    ELSIF ((x0 = TRUE) AND  (t0.Q = TRUE) AND  (t1.Q = FALSE)) THEN 
        cstate16 := 38115; y0 := TRUE; y1 := FALSE; y2 := FALSE; t0_start := TRUE; t0_up := FALSE;t1_start := FALSE; 
    ELSIF ((x0 = TRUE) AND  (t0.Q = TRUE) AND  (t1.Q = TRUE)) THEN 
        cstate16 := 39140; y0 := TRUE; y1 := FALSE; y2 := FALSE; t0_start := TRUE; t0_up := FALSE;t1_start := FALSE; 
    END_IF;
42457:
    IF ((x0 = FALSE) AND  (t0.Q = FALSE) AND  (t1.Q = FALSE)) THEN 
        cstate16 := 32883; y0 := FALSE; y1 := FALSE; y2 := FALSE; t0_start := FALSE;t1_start := FALSE; 
    ELSIF ((x0 = FALSE) AND  (t0.Q = FALSE) AND  (t1.Q = TRUE)) THEN 
        cstate16 := 34932; y0 := FALSE; y1 := FALSE; y2 := FALSE; t0_start := FALSE;t1_start := FALSE; 
    ELSIF ((x0 = FALSE) AND  (t0.Q = TRUE) AND  (t1.Q = FALSE)) THEN 
        cstate16 := 27763; y0 := FALSE; y1 := FALSE; y2 := FALSE; t0_start := FALSE;t1_start := FALSE; 
    ELSIF ((x0 = FALSE) AND  (t0.Q = TRUE) AND  (t1.Q = TRUE)) THEN 
        cstate16 := 28788; y0 := FALSE; y1 := FALSE; y2 := FALSE; t0_start := FALSE;t1_start := FALSE; 
    ELSIF ((x0 = TRUE) AND  (t0.Q = FALSE) AND  (t1.Q = FALSE)) THEN 
        cstate16 := 49657; y0 := TRUE; y1 := TRUE; y2 := TRUE; t0_start := FALSE;t1_start := FALSE; 
    ELSIF ((x0 = TRUE) AND  (t0.Q = FALSE) AND  (t1.Q = TRUE)) THEN 
        cstate16 := 48646; y0 := TRUE; y1 := TRUE; y2 := TRUE; t0_start := FALSE;t1_start := FALSE; 
    ELSIF ((x0 = TRUE) AND  (t0.Q = TRUE) AND  (t1.Q = FALSE)) THEN 
        cstate16 := 42489; y0 := TRUE; y1 := TRUE; y2 := TRUE; t0_start := FALSE;t1_start := FALSE; 
    ELSIF ((x0 = TRUE) AND  (t0.Q = TRUE) AND  (t1.Q = TRUE)) THEN 
        cstate16 := 43526; y0 := TRUE; y1 := TRUE; y2 := TRUE; t0_start := FALSE;t1_start := FALSE; 
    END_IF;
27731:
    IF ((x0 = FALSE) AND  (t0.Q = FALSE) AND  (t1.Q = FALSE)) THEN 
        cstate16 := 32883; y0 := FALSE; y1 := FALSE; y2 := FALSE; t0_start := FALSE;t1_start := FALSE; 
    ELSIF ((x0 = FALSE) AND  (t0.Q = FALSE) AND  (t1.Q = TRUE)) THEN 
        cstate16 := 34932; y0 := FALSE; y1 := FALSE; y2 := FALSE; t0_start := FALSE;t1_start := FALSE; 
    ELSIF ((x0 = FALSE) AND  (t0.Q = TRUE) AND  (t1.Q = FALSE)) THEN 
        cstate16 := 27763; y0 := FALSE; y1 := FALSE; y2 := FALSE; t0_start := FALSE;t1_start := FALSE; 
    ELSIF ((x0 = FALSE) AND  (t0.Q = TRUE) AND  (t1.Q = TRUE)) THEN 
        cstate16 := 28788; y0 := FALSE; y1 := FALSE; y2 := FALSE; t0_start := FALSE;t1_start := FALSE; 
    ELSIF ((x0 = TRUE) AND  (t0.Q = FALSE) AND  (t1.Q = FALSE)) THEN 
        cstate16 := 41187; y0 := TRUE; y1 := FALSE; y2 := FALSE; t0_start := TRUE; t0_up := FALSE;t1_start := FALSE; 
    ELSIF ((x0 = TRUE) AND  (t0.Q = FALSE) AND  (t1.Q = TRUE)) THEN 
        cstate16 := 40167; y0 := TRUE; y1 := FALSE; y2 := TRUE; t0_start := TRUE; t0_up := FALSE;t1_start := FALSE; 
    ELSIF ((x0 = TRUE) AND  (t0.Q = TRUE) AND  (t1.Q = FALSE)) THEN 
        cstate16 := 38115; y0 := TRUE; y1 := FALSE; y2 := FALSE; t0_start := TRUE; t0_up := FALSE;t1_start := FALSE; 
    ELSIF ((x0 = TRUE) AND  (t0.Q = TRUE) AND  (t1.Q = TRUE)) THEN 
        cstate16 := 39143; y0 := TRUE; y1 := FALSE; y2 := TRUE; t0_start := TRUE; t0_up := FALSE;t1_start := FALSE; 
    END_IF;
41555:
    IF ((x0 = FALSE) AND  (t0.Q = FALSE) AND  (t1.Q = FALSE)) THEN 
        cstate16 := 23667; y0 := FALSE; y1 := FALSE; y2 := FALSE; t0_start := FALSE;t1_start := FALSE; 
    ELSIF ((x0 = FALSE) AND  (t0.Q = FALSE) AND  (t1.Q = TRUE)) THEN 
        cstate16 := 26740; y0 := FALSE; y1 := FALSE; y2 := FALSE; t0_start := FALSE;t1_start := FALSE; 
    ELSIF ((x0 = FALSE) AND  (t0.Q = TRUE) AND  (t1.Q = FALSE)) THEN 
        cstate16 := 17491; y0 := FALSE; y1 := FALSE; y2 := FALSE; t0_start := FALSE;t1_start := TRUE; t1_up := FALSE; 
    ELSIF ((x0 = FALSE) AND  (t0.Q = TRUE) AND  (t1.Q = TRUE)) THEN 
        cstate16 := 17492; y0 := FALSE; y1 := FALSE; y2 := FALSE; t0_start := FALSE;t1_start := TRUE; t1_up := FALSE; 
    ELSIF ((x0 = TRUE) AND  (t0.Q = FALSE) AND  (t1.Q = FALSE)) THEN 
        cstate16 := 41555; y0 := TRUE; y1 := FALSE; y2 := FALSE; t0_start := FALSE;t1_start := FALSE; 
    ELSIF ((x0 = TRUE) AND  (t0.Q = FALSE) AND  (t1.Q = TRUE)) THEN 
        cstate16 := 40535; y0 := TRUE; y1 := FALSE; y2 := TRUE; t0_start := FALSE;t1_start := FALSE; 
    ELSIF ((x0 = TRUE) AND  (t0.Q = TRUE) AND  (t1.Q = FALSE)) THEN 
        cstate16 := 46643; y0 := TRUE; y1 := TRUE; y2 := FALSE; t0_start := FALSE;t1_start := TRUE; t1_up := FALSE; 
    ELSIF ((x0 = TRUE) AND  (t0.Q = TRUE) AND  (t1.Q = TRUE)) THEN 
        cstate16 := 46648; y0 := TRUE; y1 := TRUE; y2 := TRUE; t0_start := FALSE;t1_start := TRUE; t1_up := FALSE; 
    END_IF;
42453:
    IF ((x0 = FALSE) AND  (t0.Q = FALSE) AND  (t1.Q = FALSE)) THEN 
        cstate16 := 32883; y0 := FALSE; y1 := FALSE; y2 := FALSE; t0_start := FALSE;t1_start := FALSE; 
    ELSIF ((x0 = FALSE) AND  (t0.Q = FALSE) AND  (t1.Q = TRUE)) THEN 
        cstate16 := 34932; y0 := FALSE; y1 := FALSE; y2 := FALSE; t0_start := FALSE;t1_start := FALSE; 
    ELSIF ((x0 = FALSE) AND  (t0.Q = TRUE) AND  (t1.Q = FALSE)) THEN 
        cstate16 := 27763; y0 := FALSE; y1 := FALSE; y2 := FALSE; t0_start := FALSE;t1_start := FALSE; 
    ELSIF ((x0 = FALSE) AND  (t0.Q = TRUE) AND  (t1.Q = TRUE)) THEN 
        cstate16 := 28788; y0 := FALSE; y1 := FALSE; y2 := FALSE; t0_start := FALSE;t1_start := FALSE; 
    ELSIF ((x0 = TRUE) AND  (t0.Q = FALSE) AND  (t1.Q = FALSE)) THEN 
        cstate16 := 49657; y0 := TRUE; y1 := TRUE; y2 := TRUE; t0_start := FALSE;t1_start := FALSE; 
    ELSIF ((x0 = TRUE) AND  (t0.Q = FALSE) AND  (t1.Q = TRUE)) THEN 
        cstate16 := 48646; y0 := TRUE; y1 := TRUE; y2 := TRUE; t0_start := FALSE;t1_start := FALSE; 
    ELSIF ((x0 = TRUE) AND  (t0.Q = TRUE) AND  (t1.Q = FALSE)) THEN 
        cstate16 := 42489; y0 := TRUE; y1 := TRUE; y2 := TRUE; t0_start := FALSE;t1_start := FALSE; 
    ELSIF ((x0 = TRUE) AND  (t0.Q = TRUE) AND  (t1.Q = TRUE)) THEN 
        cstate16 := 43526; y0 := TRUE; y1 := TRUE; y2 := TRUE; t0_start := FALSE;t1_start := FALSE; 
    END_IF;
42450:
    IF ((x0 = FALSE) AND  (t0.Q = FALSE) AND  (t1.Q = FALSE)) THEN 
        cstate16 := 32883; y0 := FALSE; y1 := FALSE; y2 := FALSE; t0_start := FALSE;t1_start := FALSE; 
    ELSIF ((x0 = FALSE) AND  (t0.Q = FALSE) AND  (t1.Q = TRUE)) THEN 
        cstate16 := 34932; y0 := FALSE; y1 := FALSE; y2 := FALSE; t0_start := FALSE;t1_start := FALSE; 
    ELSIF ((x0 = FALSE) AND  (t0.Q = TRUE) AND  (t1.Q = FALSE)) THEN 
        cstate16 := 27763; y0 := FALSE; y1 := FALSE; y2 := FALSE; t0_start := FALSE;t1_start := FALSE; 
    ELSIF ((x0 = FALSE) AND  (t0.Q = TRUE) AND  (t1.Q = TRUE)) THEN 
        cstate16 := 28788; y0 := FALSE; y1 := FALSE; y2 := FALSE; t0_start := FALSE;t1_start := FALSE; 
    ELSIF ((x0 = TRUE) AND  (t0.Q = FALSE) AND  (t1.Q = FALSE)) THEN 
        cstate16 := 49649; y0 := TRUE; y1 := TRUE; y2 := FALSE; t0_start := FALSE;t1_start := FALSE; 
    ELSIF ((x0 = TRUE) AND  (t0.Q = FALSE) AND  (t1.Q = TRUE)) THEN 
        cstate16 := 48642; y0 := TRUE; y1 := TRUE; y2 := FALSE; t0_start := FALSE;t1_start := FALSE; 
    ELSIF ((x0 = TRUE) AND  (t0.Q = TRUE) AND  (t1.Q = FALSE)) THEN 
        cstate16 := 42481; y0 := TRUE; y1 := TRUE; y2 := FALSE; t0_start := FALSE;t1_start := FALSE; 
    ELSIF ((x0 = TRUE) AND  (t0.Q = TRUE) AND  (t1.Q = TRUE)) THEN 
        cstate16 := 43522; y0 := TRUE; y1 := TRUE; y2 := FALSE; t0_start := FALSE;t1_start := FALSE; 
    END_IF;
26740:
    IF ((x0 = FALSE) AND  (t0.Q = FALSE) AND  (t1.Q = FALSE)) THEN 
        cstate16 := 26739; y0 := FALSE; y1 := FALSE; y2 := FALSE; t0_start := FALSE;t1_start := FALSE; 
    ELSIF ((x0 = FALSE) AND  (t0.Q = FALSE) AND  (t1.Q = TRUE)) THEN 
        cstate16 := 26740; y0 := FALSE; y1 := FALSE; y2 := FALSE; t0_start := FALSE;t1_start := FALSE; 
    ELSIF ((x0 = FALSE) AND  (t0.Q = TRUE) AND  (t1.Q = FALSE)) THEN 
        cstate16 := 17491; y0 := FALSE; y1 := FALSE; y2 := FALSE; t0_start := FALSE;t1_start := TRUE; t1_up := FALSE; 
    ELSIF ((x0 = FALSE) AND  (t0.Q = TRUE) AND  (t1.Q = TRUE)) THEN 
        cstate16 := 17492; y0 := FALSE; y1 := FALSE; y2 := FALSE; t0_start := FALSE;t1_start := TRUE; t1_up := FALSE; 
    ELSIF ((x0 = TRUE) AND  (t0.Q = FALSE) AND  (t1.Q = FALSE)) THEN 
        cstate16 := 40163; y0 := TRUE; y1 := FALSE; y2 := FALSE; t0_start := TRUE; t0_up := FALSE;t1_start := FALSE; 
    ELSIF ((x0 = TRUE) AND  (t0.Q = FALSE) AND  (t1.Q = TRUE)) THEN 
        cstate16 := 40164; y0 := TRUE; y1 := FALSE; y2 := FALSE; t0_start := TRUE; t0_up := FALSE;t1_start := FALSE; 
    ELSIF ((x0 = TRUE) AND  (t0.Q = TRUE) AND  (t1.Q = FALSE)) THEN 
        cstate16 := 38147; y0 := TRUE; y1 := TRUE; y2 := FALSE; t0_start := TRUE; t0_up := FALSE;t1_start := TRUE; t1_up := FALSE; 
    ELSIF ((x0 = TRUE) AND  (t0.Q = TRUE) AND  (t1.Q = TRUE)) THEN 
        cstate16 := 38148; y0 := TRUE; y1 := TRUE; y2 := FALSE; t0_start := TRUE; t0_up := FALSE;t1_start := TRUE; t1_up := FALSE; 
    END_IF;
40532:
    IF ((x0 = FALSE) AND  (t0.Q = FALSE) AND  (t1.Q = FALSE)) THEN 
        cstate16 := 26739; y0 := FALSE; y1 := FALSE; y2 := FALSE; t0_start := FALSE;t1_start := FALSE; 
    ELSIF ((x0 = FALSE) AND  (t0.Q = FALSE) AND  (t1.Q = TRUE)) THEN 
        cstate16 := 26740; y0 := FALSE; y1 := FALSE; y2 := FALSE; t0_start := FALSE;t1_start := FALSE; 
    ELSIF ((x0 = FALSE) AND  (t0.Q = TRUE) AND  (t1.Q = FALSE)) THEN 
        cstate16 := 17491; y0 := FALSE; y1 := FALSE; y2 := FALSE; t0_start := FALSE;t1_start := TRUE; t1_up := FALSE; 
    ELSIF ((x0 = FALSE) AND  (t0.Q = TRUE) AND  (t1.Q = TRUE)) THEN 
        cstate16 := 17492; y0 := FALSE; y1 := FALSE; y2 := FALSE; t0_start := FALSE;t1_start := TRUE; t1_up := FALSE; 
    ELSIF ((x0 = TRUE) AND  (t0.Q = FALSE) AND  (t1.Q = FALSE)) THEN 
        cstate16 := 40531; y0 := TRUE; y1 := FALSE; y2 := FALSE; t0_start := FALSE;t1_start := FALSE; 
    ELSIF ((x0 = TRUE) AND  (t0.Q = FALSE) AND  (t1.Q = TRUE)) THEN 
        cstate16 := 40532; y0 := TRUE; y1 := FALSE; y2 := FALSE; t0_start := FALSE;t1_start := FALSE; 
    ELSIF ((x0 = TRUE) AND  (t0.Q = TRUE) AND  (t1.Q = FALSE)) THEN 
        cstate16 := 46643; y0 := TRUE; y1 := TRUE; y2 := FALSE; t0_start := FALSE;t1_start := TRUE; t1_up := FALSE; 
    ELSIF ((x0 = TRUE) AND  (t0.Q = TRUE) AND  (t1.Q = TRUE)) THEN 
        cstate16 := 46644; y0 := TRUE; y1 := TRUE; y2 := FALSE; t0_start := FALSE;t1_start := TRUE; t1_up := FALSE; 
    END_IF;
40535:
    IF ((x0 = FALSE) AND  (t0.Q = FALSE) AND  (t1.Q = FALSE)) THEN 
        cstate16 := 26739; y0 := FALSE; y1 := FALSE; y2 := FALSE; t0_start := FALSE;t1_start := FALSE; 
    ELSIF ((x0 = FALSE) AND  (t0.Q = FALSE) AND  (t1.Q = TRUE)) THEN 
        cstate16 := 26740; y0 := FALSE; y1 := FALSE; y2 := FALSE; t0_start := FALSE;t1_start := FALSE; 
    ELSIF ((x0 = FALSE) AND  (t0.Q = TRUE) AND  (t1.Q = FALSE)) THEN 
        cstate16 := 17491; y0 := FALSE; y1 := FALSE; y2 := FALSE; t0_start := FALSE;t1_start := TRUE; t1_up := FALSE; 
    ELSIF ((x0 = FALSE) AND  (t0.Q = TRUE) AND  (t1.Q = TRUE)) THEN 
        cstate16 := 17492; y0 := FALSE; y1 := FALSE; y2 := FALSE; t0_start := FALSE;t1_start := TRUE; t1_up := FALSE; 
    ELSIF ((x0 = TRUE) AND  (t0.Q = FALSE) AND  (t1.Q = FALSE)) THEN 
        cstate16 := 40540; y0 := TRUE; y1 := FALSE; y2 := TRUE; t0_start := FALSE;t1_start := FALSE; 
    ELSIF ((x0 = TRUE) AND  (t0.Q = FALSE) AND  (t1.Q = TRUE)) THEN 
        cstate16 := 40535; y0 := TRUE; y1 := FALSE; y2 := TRUE; t0_start := FALSE;t1_start := FALSE; 
    ELSIF ((x0 = TRUE) AND  (t0.Q = TRUE) AND  (t1.Q = FALSE)) THEN 
        cstate16 := 46651; y0 := TRUE; y1 := TRUE; y2 := TRUE; t0_start := FALSE;t1_start := TRUE; t1_up := FALSE; 
    ELSIF ((x0 = TRUE) AND  (t0.Q = TRUE) AND  (t1.Q = TRUE)) THEN 
        cstate16 := 46648; y0 := TRUE; y1 := TRUE; y2 := TRUE; t0_start := FALSE;t1_start := TRUE; t1_up := FALSE; 
    END_IF;
6481:
    IF ((x0 = FALSE) AND  (t0.Q = FALSE) AND  (t1.Q = FALSE)) THEN 
        cstate16 := 34931; y0 := FALSE; y1 := FALSE; y2 := FALSE; t0_start := FALSE;t1_start := FALSE; 
    ELSIF ((x0 = FALSE) AND  (t0.Q = FALSE) AND  (t1.Q = TRUE)) THEN 
        cstate16 := 34932; y0 := FALSE; y1 := FALSE; y2 := FALSE; t0_start := FALSE;t1_start := FALSE; 
    ELSIF ((x0 = FALSE) AND  (t0.Q = TRUE) AND  (t1.Q = FALSE)) THEN 
        cstate16 := 28787; y0 := FALSE; y1 := FALSE; y2 := FALSE; t0_start := FALSE;t1_start := FALSE; 
    ELSIF ((x0 = FALSE) AND  (t0.Q = TRUE) AND  (t1.Q = TRUE)) THEN 
        cstate16 := 28788; y0 := FALSE; y1 := FALSE; y2 := FALSE; t0_start := FALSE;t1_start := FALSE; 
    ELSIF ((x0 = TRUE) AND  (t0.Q = FALSE) AND  (t1.Q = FALSE)) THEN 
        cstate16 := 14673; y0 := FALSE; y1 := TRUE; y2 := FALSE; t0_start := FALSE;t1_start := FALSE; 
    ELSIF ((x0 = TRUE) AND  (t0.Q = FALSE) AND  (t1.Q = TRUE)) THEN 
        cstate16 := 14678; y0 := FALSE; y1 := TRUE; y2 := TRUE; t0_start := FALSE;t1_start := FALSE; 
    ELSIF ((x0 = TRUE) AND  (t0.Q = TRUE) AND  (t1.Q = FALSE)) THEN 
        cstate16 := 6481; y0 := FALSE; y1 := TRUE; y2 := FALSE; t0_start := FALSE;t1_start := FALSE; 
    ELSIF ((x0 = TRUE) AND  (t0.Q = TRUE) AND  (t1.Q = TRUE)) THEN 
        cstate16 := 6486; y0 := FALSE; y1 := TRUE; y2 := TRUE; t0_start := FALSE;t1_start := FALSE; 
    END_IF;
6482:
    IF ((x0 = FALSE) AND  (t0.Q = FALSE) AND  (t1.Q = FALSE)) THEN 
        cstate16 := 34931; y0 := FALSE; y1 := FALSE; y2 := FALSE; t0_start := FALSE;t1_start := FALSE; 
    ELSIF ((x0 = FALSE) AND  (t0.Q = FALSE) AND  (t1.Q = TRUE)) THEN 
        cstate16 := 34932; y0 := FALSE; y1 := FALSE; y2 := FALSE; t0_start := FALSE;t1_start := FALSE; 
    ELSIF ((x0 = FALSE) AND  (t0.Q = TRUE) AND  (t1.Q = FALSE)) THEN 
        cstate16 := 28787; y0 := FALSE; y1 := FALSE; y2 := FALSE; t0_start := FALSE;t1_start := FALSE; 
    ELSIF ((x0 = FALSE) AND  (t0.Q = TRUE) AND  (t1.Q = TRUE)) THEN 
        cstate16 := 28788; y0 := FALSE; y1 := FALSE; y2 := FALSE; t0_start := FALSE;t1_start := FALSE; 
    ELSIF ((x0 = TRUE) AND  (t0.Q = FALSE) AND  (t1.Q = FALSE)) THEN 
        cstate16 := 14673; y0 := FALSE; y1 := TRUE; y2 := FALSE; t0_start := FALSE;t1_start := FALSE; 
    ELSIF ((x0 = TRUE) AND  (t0.Q = FALSE) AND  (t1.Q = TRUE)) THEN 
        cstate16 := 14674; y0 := FALSE; y1 := TRUE; y2 := FALSE; t0_start := FALSE;t1_start := FALSE; 
    ELSIF ((x0 = TRUE) AND  (t0.Q = TRUE) AND  (t1.Q = FALSE)) THEN 
        cstate16 := 6481; y0 := FALSE; y1 := TRUE; y2 := FALSE; t0_start := FALSE;t1_start := FALSE; 
    ELSIF ((x0 = TRUE) AND  (t0.Q = TRUE) AND  (t1.Q = TRUE)) THEN 
        cstate16 := 6482; y0 := FALSE; y1 := TRUE; y2 := FALSE; t0_start := FALSE;t1_start := FALSE; 
    END_IF;
26138:
    IF ((x0 = FALSE) AND  (t0.Q = FALSE) AND  (t1.Q = FALSE)) THEN 
        cstate16 := 26739; y0 := FALSE; y1 := FALSE; y2 := FALSE; t0_start := FALSE;t1_start := FALSE; 
    ELSIF ((x0 = FALSE) AND  (t0.Q = FALSE) AND  (t1.Q = TRUE)) THEN 
        cstate16 := 26740; y0 := FALSE; y1 := FALSE; y2 := FALSE; t0_start := FALSE;t1_start := FALSE; 
    ELSIF ((x0 = FALSE) AND  (t0.Q = TRUE) AND  (t1.Q = FALSE)) THEN 
        cstate16 := 17491; y0 := FALSE; y1 := FALSE; y2 := FALSE; t0_start := FALSE;t1_start := TRUE; t1_up := FALSE; 
    ELSIF ((x0 = FALSE) AND  (t0.Q = TRUE) AND  (t1.Q = TRUE)) THEN 
        cstate16 := 17492; y0 := FALSE; y1 := FALSE; y2 := FALSE; t0_start := FALSE;t1_start := TRUE; t1_up := FALSE; 
    ELSIF ((x0 = TRUE) AND  (t0.Q = FALSE) AND  (t1.Q = FALSE)) THEN 
        cstate16 := 26138; y0 := TRUE; y1 := TRUE; y2 := TRUE; t0_start := FALSE;t1_start := FALSE; 
    ELSIF ((x0 = TRUE) AND  (t0.Q = FALSE) AND  (t1.Q = TRUE)) THEN 
        cstate16 := 26134; y0 := TRUE; y1 := TRUE; y2 := TRUE; t0_start := FALSE;t1_start := FALSE; 
    ELSIF ((x0 = TRUE) AND  (t0.Q = TRUE) AND  (t1.Q = FALSE)) THEN 
        cstate16 := 42457; y0 := TRUE; y1 := TRUE; y2 := TRUE; t0_start := FALSE;t1_start := TRUE; t1_up := FALSE; 
    ELSIF ((x0 = TRUE) AND  (t0.Q = TRUE) AND  (t1.Q = TRUE)) THEN 
        cstate16 := 42453; y0 := TRUE; y1 := TRUE; y2 := TRUE; t0_start := FALSE;t1_start := TRUE; t1_up := FALSE; 
    END_IF;
6486:
    IF ((x0 = FALSE) AND  (t0.Q = FALSE) AND  (t1.Q = FALSE)) THEN 
        cstate16 := 34931; y0 := FALSE; y1 := FALSE; y2 := FALSE; t0_start := FALSE;t1_start := FALSE; 
    ELSIF ((x0 = FALSE) AND  (t0.Q = FALSE) AND  (t1.Q = TRUE)) THEN 
        cstate16 := 34932; y0 := FALSE; y1 := FALSE; y2 := FALSE; t0_start := FALSE;t1_start := FALSE; 
    ELSIF ((x0 = FALSE) AND  (t0.Q = TRUE) AND  (t1.Q = FALSE)) THEN 
        cstate16 := 28787; y0 := FALSE; y1 := FALSE; y2 := FALSE; t0_start := FALSE;t1_start := FALSE; 
    ELSIF ((x0 = FALSE) AND  (t0.Q = TRUE) AND  (t1.Q = TRUE)) THEN 
        cstate16 := 28788; y0 := FALSE; y1 := FALSE; y2 := FALSE; t0_start := FALSE;t1_start := FALSE; 
    ELSIF ((x0 = TRUE) AND  (t0.Q = FALSE) AND  (t1.Q = FALSE)) THEN 
        cstate16 := 14682; y0 := FALSE; y1 := TRUE; y2 := TRUE; t0_start := FALSE;t1_start := FALSE; 
    ELSIF ((x0 = TRUE) AND  (t0.Q = FALSE) AND  (t1.Q = TRUE)) THEN 
        cstate16 := 14678; y0 := FALSE; y1 := TRUE; y2 := TRUE; t0_start := FALSE;t1_start := FALSE; 
    ELSIF ((x0 = TRUE) AND  (t0.Q = TRUE) AND  (t1.Q = FALSE)) THEN 
        cstate16 := 6490; y0 := FALSE; y1 := TRUE; y2 := TRUE; t0_start := FALSE;t1_start := FALSE; 
    ELSIF ((x0 = TRUE) AND  (t0.Q = TRUE) AND  (t1.Q = TRUE)) THEN 
        cstate16 := 6486; y0 := FALSE; y1 := TRUE; y2 := TRUE; t0_start := FALSE;t1_start := FALSE; 
    END_IF;
40531:
    IF ((x0 = FALSE) AND  (t0.Q = FALSE) AND  (t1.Q = FALSE)) THEN 
        cstate16 := 26739; y0 := FALSE; y1 := FALSE; y2 := FALSE; t0_start := FALSE;t1_start := FALSE; 
    ELSIF ((x0 = FALSE) AND  (t0.Q = FALSE) AND  (t1.Q = TRUE)) THEN 
        cstate16 := 26740; y0 := FALSE; y1 := FALSE; y2 := FALSE; t0_start := FALSE;t1_start := FALSE; 
    ELSIF ((x0 = FALSE) AND  (t0.Q = TRUE) AND  (t1.Q = FALSE)) THEN 
        cstate16 := 17491; y0 := FALSE; y1 := FALSE; y2 := FALSE; t0_start := FALSE;t1_start := TRUE; t1_up := FALSE; 
    ELSIF ((x0 = FALSE) AND  (t0.Q = TRUE) AND  (t1.Q = TRUE)) THEN 
        cstate16 := 17492; y0 := FALSE; y1 := FALSE; y2 := FALSE; t0_start := FALSE;t1_start := TRUE; t1_up := FALSE; 
    ELSIF ((x0 = TRUE) AND  (t0.Q = FALSE) AND  (t1.Q = FALSE)) THEN 
        cstate16 := 40531; y0 := TRUE; y1 := FALSE; y2 := FALSE; t0_start := FALSE;t1_start := FALSE; 
    ELSIF ((x0 = TRUE) AND  (t0.Q = FALSE) AND  (t1.Q = TRUE)) THEN 
        cstate16 := 40535; y0 := TRUE; y1 := FALSE; y2 := TRUE; t0_start := FALSE;t1_start := FALSE; 
    ELSIF ((x0 = TRUE) AND  (t0.Q = TRUE) AND  (t1.Q = FALSE)) THEN 
        cstate16 := 46643; y0 := TRUE; y1 := TRUE; y2 := FALSE; t0_start := FALSE;t1_start := TRUE; t1_up := FALSE; 
    ELSIF ((x0 = TRUE) AND  (t0.Q = TRUE) AND  (t1.Q = TRUE)) THEN 
        cstate16 := 46648; y0 := TRUE; y1 := TRUE; y2 := TRUE; t0_start := FALSE;t1_start := TRUE; t1_up := FALSE; 
    END_IF;
39140:
    IF ((x0 = FALSE) AND  (t0.Q = FALSE) AND  (t1.Q = FALSE)) THEN 
        cstate16 := 26739; y0 := FALSE; y1 := FALSE; y2 := FALSE; t0_start := FALSE;t1_start := FALSE; 
    ELSIF ((x0 = FALSE) AND  (t0.Q = FALSE) AND  (t1.Q = TRUE)) THEN 
        cstate16 := 26740; y0 := FALSE; y1 := FALSE; y2 := FALSE; t0_start := FALSE;t1_start := FALSE; 
    ELSIF ((x0 = FALSE) AND  (t0.Q = TRUE) AND  (t1.Q = FALSE)) THEN 
        cstate16 := 22643; y0 := FALSE; y1 := FALSE; y2 := FALSE; t0_start := FALSE;t1_start := FALSE; 
    ELSIF ((x0 = FALSE) AND  (t0.Q = TRUE) AND  (t1.Q = TRUE)) THEN 
        cstate16 := 22644; y0 := FALSE; y1 := FALSE; y2 := FALSE; t0_start := FALSE;t1_start := FALSE; 
    ELSIF ((x0 = TRUE) AND  (t0.Q = FALSE) AND  (t1.Q = FALSE)) THEN 
        cstate16 := 40531; y0 := TRUE; y1 := FALSE; y2 := FALSE; t0_start := FALSE;t1_start := FALSE; 
    ELSIF ((x0 = TRUE) AND  (t0.Q = FALSE) AND  (t1.Q = TRUE)) THEN 
        cstate16 := 40532; y0 := TRUE; y1 := FALSE; y2 := FALSE; t0_start := FALSE;t1_start := FALSE; 
    ELSIF ((x0 = TRUE) AND  (t0.Q = TRUE) AND  (t1.Q = FALSE)) THEN 
        cstate16 := 47683; y0 := TRUE; y1 := FALSE; y2 := FALSE; t0_start := FALSE;t1_start := FALSE; 
    ELSIF ((x0 = TRUE) AND  (t0.Q = TRUE) AND  (t1.Q = TRUE)) THEN 
        cstate16 := 47684; y0 := TRUE; y1 := FALSE; y2 := FALSE; t0_start := FALSE;t1_start := FALSE; 
    END_IF;
40663:
    IF ((x0 = FALSE) AND  (t0.Q = FALSE) AND  (t1.Q = FALSE)) THEN 
        cstate16 := 26739; y0 := FALSE; y1 := FALSE; y2 := FALSE; t0_start := FALSE;t1_start := FALSE; 
    ELSIF ((x0 = FALSE) AND  (t0.Q = FALSE) AND  (t1.Q = TRUE)) THEN 
        cstate16 := 26740; y0 := FALSE; y1 := FALSE; y2 := FALSE; t0_start := FALSE;t1_start := FALSE; 
    ELSIF ((x0 = FALSE) AND  (t0.Q = TRUE) AND  (t1.Q = FALSE)) THEN 
        cstate16 := 17491; y0 := FALSE; y1 := FALSE; y2 := FALSE; t0_start := FALSE;t1_start := TRUE; t1_up := FALSE; 
    ELSIF ((x0 = FALSE) AND  (t0.Q = TRUE) AND  (t1.Q = TRUE)) THEN 
        cstate16 := 17492; y0 := FALSE; y1 := FALSE; y2 := FALSE; t0_start := FALSE;t1_start := TRUE; t1_up := FALSE; 
    ELSIF ((x0 = TRUE) AND  (t0.Q = FALSE) AND  (t1.Q = FALSE)) THEN 
        cstate16 := 40668; y0 := TRUE; y1 := TRUE; y2 := TRUE; t0_start := FALSE;t1_start := FALSE; 
    ELSIF ((x0 = TRUE) AND  (t0.Q = FALSE) AND  (t1.Q = TRUE)) THEN 
        cstate16 := 40663; y0 := TRUE; y1 := TRUE; y2 := TRUE; t0_start := FALSE;t1_start := FALSE; 
    ELSIF ((x0 = TRUE) AND  (t0.Q = TRUE) AND  (t1.Q = FALSE)) THEN 
        cstate16 := 46651; y0 := TRUE; y1 := TRUE; y2 := TRUE; t0_start := FALSE;t1_start := TRUE; t1_up := FALSE; 
    ELSIF ((x0 = TRUE) AND  (t0.Q = TRUE) AND  (t1.Q = TRUE)) THEN 
        cstate16 := 46648; y0 := TRUE; y1 := TRUE; y2 := TRUE; t0_start := FALSE;t1_start := TRUE; t1_up := FALSE; 
    END_IF;
26038:
    IF ((x0 = FALSE) AND  (t0.Q = FALSE) AND  (t1.Q = FALSE)) THEN 
        cstate16 := 26739; y0 := FALSE; y1 := FALSE; y2 := FALSE; t0_start := FALSE;t1_start := FALSE; 
    ELSIF ((x0 = FALSE) AND  (t0.Q = FALSE) AND  (t1.Q = TRUE)) THEN 
        cstate16 := 26740; y0 := FALSE; y1 := FALSE; y2 := FALSE; t0_start := FALSE;t1_start := FALSE; 
    ELSIF ((x0 = FALSE) AND  (t0.Q = TRUE) AND  (t1.Q = FALSE)) THEN 
        cstate16 := 17491; y0 := FALSE; y1 := FALSE; y2 := FALSE; t0_start := FALSE;t1_start := TRUE; t1_up := FALSE; 
    ELSIF ((x0 = FALSE) AND  (t0.Q = TRUE) AND  (t1.Q = TRUE)) THEN 
        cstate16 := 17492; y0 := FALSE; y1 := FALSE; y2 := FALSE; t0_start := FALSE;t1_start := TRUE; t1_up := FALSE; 
    ELSIF ((x0 = TRUE) AND  (t0.Q = FALSE) AND  (t1.Q = FALSE)) THEN 
        cstate16 := 26042; y0 := TRUE; y1 := FALSE; y2 := TRUE; t0_start := FALSE;t1_start := FALSE; 
    ELSIF ((x0 = TRUE) AND  (t0.Q = FALSE) AND  (t1.Q = TRUE)) THEN 
        cstate16 := 26038; y0 := TRUE; y1 := FALSE; y2 := TRUE; t0_start := FALSE;t1_start := FALSE; 
    ELSIF ((x0 = TRUE) AND  (t0.Q = TRUE) AND  (t1.Q = FALSE)) THEN 
        cstate16 := 42457; y0 := TRUE; y1 := TRUE; y2 := TRUE; t0_start := FALSE;t1_start := TRUE; t1_up := FALSE; 
    ELSIF ((x0 = TRUE) AND  (t0.Q = TRUE) AND  (t1.Q = TRUE)) THEN 
        cstate16 := 42453; y0 := TRUE; y1 := TRUE; y2 := TRUE; t0_start := FALSE;t1_start := TRUE; t1_up := FALSE; 
    END_IF;
40660:
    IF ((x0 = FALSE) AND  (t0.Q = FALSE) AND  (t1.Q = FALSE)) THEN 
        cstate16 := 26739; y0 := FALSE; y1 := FALSE; y2 := FALSE; t0_start := FALSE;t1_start := FALSE; 
    ELSIF ((x0 = FALSE) AND  (t0.Q = FALSE) AND  (t1.Q = TRUE)) THEN 
        cstate16 := 26740; y0 := FALSE; y1 := FALSE; y2 := FALSE; t0_start := FALSE;t1_start := FALSE; 
    ELSIF ((x0 = FALSE) AND  (t0.Q = TRUE) AND  (t1.Q = FALSE)) THEN 
        cstate16 := 17491; y0 := FALSE; y1 := FALSE; y2 := FALSE; t0_start := FALSE;t1_start := TRUE; t1_up := FALSE; 
    ELSIF ((x0 = FALSE) AND  (t0.Q = TRUE) AND  (t1.Q = TRUE)) THEN 
        cstate16 := 17492; y0 := FALSE; y1 := FALSE; y2 := FALSE; t0_start := FALSE;t1_start := TRUE; t1_up := FALSE; 
    ELSIF ((x0 = TRUE) AND  (t0.Q = FALSE) AND  (t1.Q = FALSE)) THEN 
        cstate16 := 40659; y0 := TRUE; y1 := TRUE; y2 := FALSE; t0_start := FALSE;t1_start := FALSE; 
    ELSIF ((x0 = TRUE) AND  (t0.Q = FALSE) AND  (t1.Q = TRUE)) THEN 
        cstate16 := 40660; y0 := TRUE; y1 := TRUE; y2 := FALSE; t0_start := FALSE;t1_start := FALSE; 
    ELSIF ((x0 = TRUE) AND  (t0.Q = TRUE) AND  (t1.Q = FALSE)) THEN 
        cstate16 := 46643; y0 := TRUE; y1 := TRUE; y2 := FALSE; t0_start := FALSE;t1_start := TRUE; t1_up := FALSE; 
    ELSIF ((x0 = TRUE) AND  (t0.Q = TRUE) AND  (t1.Q = TRUE)) THEN 
        cstate16 := 46644; y0 := TRUE; y1 := TRUE; y2 := FALSE; t0_start := FALSE;t1_start := TRUE; t1_up := FALSE; 
    END_IF;
42449:
    IF ((x0 = FALSE) AND  (t0.Q = FALSE) AND  (t1.Q = FALSE)) THEN 
        cstate16 := 32883; y0 := FALSE; y1 := FALSE; y2 := FALSE; t0_start := FALSE;t1_start := FALSE; 
    ELSIF ((x0 = FALSE) AND  (t0.Q = FALSE) AND  (t1.Q = TRUE)) THEN 
        cstate16 := 34932; y0 := FALSE; y1 := FALSE; y2 := FALSE; t0_start := FALSE;t1_start := FALSE; 
    ELSIF ((x0 = FALSE) AND  (t0.Q = TRUE) AND  (t1.Q = FALSE)) THEN 
        cstate16 := 27763; y0 := FALSE; y1 := FALSE; y2 := FALSE; t0_start := FALSE;t1_start := FALSE; 
    ELSIF ((x0 = FALSE) AND  (t0.Q = TRUE) AND  (t1.Q = TRUE)) THEN 
        cstate16 := 28788; y0 := FALSE; y1 := FALSE; y2 := FALSE; t0_start := FALSE;t1_start := FALSE; 
    ELSIF ((x0 = TRUE) AND  (t0.Q = FALSE) AND  (t1.Q = FALSE)) THEN 
        cstate16 := 49649; y0 := TRUE; y1 := TRUE; y2 := FALSE; t0_start := FALSE;t1_start := FALSE; 
    ELSIF ((x0 = TRUE) AND  (t0.Q = FALSE) AND  (t1.Q = TRUE)) THEN 
        cstate16 := 48646; y0 := TRUE; y1 := TRUE; y2 := TRUE; t0_start := FALSE;t1_start := FALSE; 
    ELSIF ((x0 = TRUE) AND  (t0.Q = TRUE) AND  (t1.Q = FALSE)) THEN 
        cstate16 := 42481; y0 := TRUE; y1 := TRUE; y2 := FALSE; t0_start := FALSE;t1_start := FALSE; 
    ELSIF ((x0 = TRUE) AND  (t0.Q = TRUE) AND  (t1.Q = TRUE)) THEN 
        cstate16 := 43526; y0 := TRUE; y1 := TRUE; y2 := TRUE; t0_start := FALSE;t1_start := FALSE; 
    END_IF;
39143:
    IF ((x0 = FALSE) AND  (t0.Q = FALSE) AND  (t1.Q = FALSE)) THEN 
        cstate16 := 26739; y0 := FALSE; y1 := FALSE; y2 := FALSE; t0_start := FALSE;t1_start := FALSE; 
    ELSIF ((x0 = FALSE) AND  (t0.Q = FALSE) AND  (t1.Q = TRUE)) THEN 
        cstate16 := 26740; y0 := FALSE; y1 := FALSE; y2 := FALSE; t0_start := FALSE;t1_start := FALSE; 
    ELSIF ((x0 = FALSE) AND  (t0.Q = TRUE) AND  (t1.Q = FALSE)) THEN 
        cstate16 := 22643; y0 := FALSE; y1 := FALSE; y2 := FALSE; t0_start := FALSE;t1_start := FALSE; 
    ELSIF ((x0 = FALSE) AND  (t0.Q = TRUE) AND  (t1.Q = TRUE)) THEN 
        cstate16 := 22644; y0 := FALSE; y1 := FALSE; y2 := FALSE; t0_start := FALSE;t1_start := FALSE; 
    ELSIF ((x0 = TRUE) AND  (t0.Q = FALSE) AND  (t1.Q = FALSE)) THEN 
        cstate16 := 40540; y0 := TRUE; y1 := FALSE; y2 := TRUE; t0_start := FALSE;t1_start := FALSE; 
    ELSIF ((x0 = TRUE) AND  (t0.Q = FALSE) AND  (t1.Q = TRUE)) THEN 
        cstate16 := 40535; y0 := TRUE; y1 := FALSE; y2 := TRUE; t0_start := FALSE;t1_start := FALSE; 
    ELSIF ((x0 = TRUE) AND  (t0.Q = TRUE) AND  (t1.Q = FALSE)) THEN 
        cstate16 := 47692; y0 := TRUE; y1 := FALSE; y2 := TRUE; t0_start := FALSE;t1_start := FALSE; 
    ELSIF ((x0 = TRUE) AND  (t0.Q = TRUE) AND  (t1.Q = TRUE)) THEN 
        cstate16 := 47687; y0 := TRUE; y1 := FALSE; y2 := TRUE; t0_start := FALSE;t1_start := FALSE; 
    END_IF;
40668:
    IF ((x0 = FALSE) AND  (t0.Q = FALSE) AND  (t1.Q = FALSE)) THEN 
        cstate16 := 26739; y0 := FALSE; y1 := FALSE; y2 := FALSE; t0_start := FALSE;t1_start := FALSE; 
    ELSIF ((x0 = FALSE) AND  (t0.Q = FALSE) AND  (t1.Q = TRUE)) THEN 
        cstate16 := 26740; y0 := FALSE; y1 := FALSE; y2 := FALSE; t0_start := FALSE;t1_start := FALSE; 
    ELSIF ((x0 = FALSE) AND  (t0.Q = TRUE) AND  (t1.Q = FALSE)) THEN 
        cstate16 := 17491; y0 := FALSE; y1 := FALSE; y2 := FALSE; t0_start := FALSE;t1_start := TRUE; t1_up := FALSE; 
    ELSIF ((x0 = FALSE) AND  (t0.Q = TRUE) AND  (t1.Q = TRUE)) THEN 
        cstate16 := 17492; y0 := FALSE; y1 := FALSE; y2 := FALSE; t0_start := FALSE;t1_start := TRUE; t1_up := FALSE; 
    ELSIF ((x0 = TRUE) AND  (t0.Q = FALSE) AND  (t1.Q = FALSE)) THEN 
        cstate16 := 40668; y0 := TRUE; y1 := TRUE; y2 := TRUE; t0_start := FALSE;t1_start := FALSE; 
    ELSIF ((x0 = TRUE) AND  (t0.Q = FALSE) AND  (t1.Q = TRUE)) THEN 
        cstate16 := 40663; y0 := TRUE; y1 := TRUE; y2 := TRUE; t0_start := FALSE;t1_start := FALSE; 
    ELSIF ((x0 = TRUE) AND  (t0.Q = TRUE) AND  (t1.Q = FALSE)) THEN 
        cstate16 := 46651; y0 := TRUE; y1 := TRUE; y2 := TRUE; t0_start := FALSE;t1_start := TRUE; t1_up := FALSE; 
    ELSIF ((x0 = TRUE) AND  (t0.Q = TRUE) AND  (t1.Q = TRUE)) THEN 
        cstate16 := 46648; y0 := TRUE; y1 := TRUE; y2 := TRUE; t0_start := FALSE;t1_start := TRUE; t1_up := FALSE; 
    END_IF;
41707:
    IF ((x0 = FALSE) AND  (t0.Q = FALSE) AND  (t1.Q = FALSE)) THEN 
        cstate16 := 23667; y0 := FALSE; y1 := FALSE; y2 := FALSE; t0_start := FALSE;t1_start := FALSE; 
    ELSIF ((x0 = FALSE) AND  (t0.Q = FALSE) AND  (t1.Q = TRUE)) THEN 
        cstate16 := 26740; y0 := FALSE; y1 := FALSE; y2 := FALSE; t0_start := FALSE;t1_start := FALSE; 
    ELSIF ((x0 = FALSE) AND  (t0.Q = TRUE) AND  (t1.Q = FALSE)) THEN 
        cstate16 := 17491; y0 := FALSE; y1 := FALSE; y2 := FALSE; t0_start := FALSE;t1_start := TRUE; t1_up := FALSE; 
    ELSIF ((x0 = FALSE) AND  (t0.Q = TRUE) AND  (t1.Q = TRUE)) THEN 
        cstate16 := 17492; y0 := FALSE; y1 := FALSE; y2 := FALSE; t0_start := FALSE;t1_start := TRUE; t1_up := FALSE; 
    ELSIF ((x0 = TRUE) AND  (t0.Q = FALSE) AND  (t1.Q = FALSE)) THEN 
        cstate16 := 41707; y0 := TRUE; y1 := TRUE; y2 := TRUE; t0_start := FALSE;t1_start := FALSE; 
    ELSIF ((x0 = TRUE) AND  (t0.Q = FALSE) AND  (t1.Q = TRUE)) THEN 
        cstate16 := 40663; y0 := TRUE; y1 := TRUE; y2 := TRUE; t0_start := FALSE;t1_start := FALSE; 
    ELSIF ((x0 = TRUE) AND  (t0.Q = TRUE) AND  (t1.Q = FALSE)) THEN 
        cstate16 := 46651; y0 := TRUE; y1 := TRUE; y2 := TRUE; t0_start := FALSE;t1_start := TRUE; t1_up := FALSE; 
    ELSIF ((x0 = TRUE) AND  (t0.Q = TRUE) AND  (t1.Q = TRUE)) THEN 
        cstate16 := 46648; y0 := TRUE; y1 := TRUE; y2 := TRUE; t0_start := FALSE;t1_start := TRUE; t1_up := FALSE; 
    END_IF;
26129:
    IF ((x0 = FALSE) AND  (t0.Q = FALSE) AND  (t1.Q = FALSE)) THEN 
        cstate16 := 26739; y0 := FALSE; y1 := FALSE; y2 := FALSE; t0_start := FALSE;t1_start := FALSE; 
    ELSIF ((x0 = FALSE) AND  (t0.Q = FALSE) AND  (t1.Q = TRUE)) THEN 
        cstate16 := 26740; y0 := FALSE; y1 := FALSE; y2 := FALSE; t0_start := FALSE;t1_start := FALSE; 
    ELSIF ((x0 = FALSE) AND  (t0.Q = TRUE) AND  (t1.Q = FALSE)) THEN 
        cstate16 := 17491; y0 := FALSE; y1 := FALSE; y2 := FALSE; t0_start := FALSE;t1_start := TRUE; t1_up := FALSE; 
    ELSIF ((x0 = FALSE) AND  (t0.Q = TRUE) AND  (t1.Q = TRUE)) THEN 
        cstate16 := 17492; y0 := FALSE; y1 := FALSE; y2 := FALSE; t0_start := FALSE;t1_start := TRUE; t1_up := FALSE; 
    ELSIF ((x0 = TRUE) AND  (t0.Q = FALSE) AND  (t1.Q = FALSE)) THEN 
        cstate16 := 26129; y0 := TRUE; y1 := TRUE; y2 := FALSE; t0_start := FALSE;t1_start := FALSE; 
    ELSIF ((x0 = TRUE) AND  (t0.Q = FALSE) AND  (t1.Q = TRUE)) THEN 
        cstate16 := 26134; y0 := TRUE; y1 := TRUE; y2 := TRUE; t0_start := FALSE;t1_start := FALSE; 
    ELSIF ((x0 = TRUE) AND  (t0.Q = TRUE) AND  (t1.Q = FALSE)) THEN 
        cstate16 := 42449; y0 := TRUE; y1 := TRUE; y2 := FALSE; t0_start := FALSE;t1_start := TRUE; t1_up := FALSE; 
    ELSIF ((x0 = TRUE) AND  (t0.Q = TRUE) AND  (t1.Q = TRUE)) THEN 
        cstate16 := 42453; y0 := TRUE; y1 := TRUE; y2 := TRUE; t0_start := FALSE;t1_start := TRUE; t1_up := FALSE; 
    END_IF;
20678:
    IF ((x0 = FALSE) AND  (t0.Q = FALSE) AND  (t1.Q = FALSE)) THEN 
        cstate16 := 26739; y0 := FALSE; y1 := FALSE; y2 := FALSE; t0_start := FALSE;t1_start := FALSE; 
    ELSIF ((x0 = FALSE) AND  (t0.Q = FALSE) AND  (t1.Q = TRUE)) THEN 
        cstate16 := 26740; y0 := FALSE; y1 := FALSE; y2 := FALSE; t0_start := FALSE;t1_start := FALSE; 
    ELSIF ((x0 = FALSE) AND  (t0.Q = TRUE) AND  (t1.Q = FALSE)) THEN 
        cstate16 := 22643; y0 := FALSE; y1 := FALSE; y2 := FALSE; t0_start := FALSE;t1_start := FALSE; 
    ELSIF ((x0 = FALSE) AND  (t0.Q = TRUE) AND  (t1.Q = TRUE)) THEN 
        cstate16 := 22644; y0 := FALSE; y1 := FALSE; y2 := FALSE; t0_start := FALSE;t1_start := FALSE; 
    ELSIF ((x0 = TRUE) AND  (t0.Q = FALSE) AND  (t1.Q = FALSE)) THEN 
        cstate16 := 26042; y0 := TRUE; y1 := FALSE; y2 := TRUE; t0_start := FALSE;t1_start := FALSE; 
    ELSIF ((x0 = TRUE) AND  (t0.Q = FALSE) AND  (t1.Q = TRUE)) THEN 
        cstate16 := 26038; y0 := TRUE; y1 := FALSE; y2 := TRUE; t0_start := FALSE;t1_start := FALSE; 
    ELSIF ((x0 = TRUE) AND  (t0.Q = TRUE) AND  (t1.Q = FALSE)) THEN 
        cstate16 := 43418; y0 := TRUE; y1 := FALSE; y2 := TRUE; t0_start := FALSE;t1_start := FALSE; 
    ELSIF ((x0 = TRUE) AND  (t0.Q = TRUE) AND  (t1.Q = TRUE)) THEN 
        cstate16 := 43414; y0 := TRUE; y1 := FALSE; y2 := TRUE; t0_start := FALSE;t1_start := FALSE; 
    END_IF;
8361:
    IF ((x0 = FALSE) AND  (t0.Q = FALSE) AND  (t1.Q = FALSE)) THEN 
        cstate16 := 32883; y0 := FALSE; y1 := FALSE; y2 := FALSE; t0_start := FALSE;t1_start := FALSE; 
    ELSIF ((x0 = FALSE) AND  (t0.Q = FALSE) AND  (t1.Q = TRUE)) THEN 
        cstate16 := 34932; y0 := FALSE; y1 := FALSE; y2 := FALSE; t0_start := FALSE;t1_start := FALSE; 
    ELSIF ((x0 = FALSE) AND  (t0.Q = TRUE) AND  (t1.Q = FALSE)) THEN 
        cstate16 := 27763; y0 := FALSE; y1 := FALSE; y2 := FALSE; t0_start := FALSE;t1_start := FALSE; 
    ELSIF ((x0 = FALSE) AND  (t0.Q = TRUE) AND  (t1.Q = TRUE)) THEN 
        cstate16 := 28788; y0 := FALSE; y1 := FALSE; y2 := FALSE; t0_start := FALSE;t1_start := FALSE; 
    ELSIF ((x0 = TRUE) AND  (t0.Q = FALSE) AND  (t1.Q = FALSE)) THEN 
        cstate16 := 16697; y0 := FALSE; y1 := TRUE; y2 := TRUE; t0_start := FALSE;t1_start := FALSE; 
    ELSIF ((x0 = TRUE) AND  (t0.Q = FALSE) AND  (t1.Q = TRUE)) THEN 
        cstate16 := 14678; y0 := FALSE; y1 := TRUE; y2 := TRUE; t0_start := FALSE;t1_start := FALSE; 
    ELSIF ((x0 = TRUE) AND  (t0.Q = TRUE) AND  (t1.Q = FALSE)) THEN 
        cstate16 := 8505; y0 := FALSE; y1 := TRUE; y2 := TRUE; t0_start := FALSE;t1_start := FALSE; 
    ELSIF ((x0 = TRUE) AND  (t0.Q = TRUE) AND  (t1.Q = TRUE)) THEN 
        cstate16 := 6486; y0 := FALSE; y1 := TRUE; y2 := TRUE; t0_start := FALSE;t1_start := FALSE; 
    END_IF;
20674:
    IF ((x0 = FALSE) AND  (t0.Q = FALSE) AND  (t1.Q = FALSE)) THEN 
        cstate16 := 26739; y0 := FALSE; y1 := FALSE; y2 := FALSE; t0_start := FALSE;t1_start := FALSE; 
    ELSIF ((x0 = FALSE) AND  (t0.Q = FALSE) AND  (t1.Q = TRUE)) THEN 
        cstate16 := 26740; y0 := FALSE; y1 := FALSE; y2 := FALSE; t0_start := FALSE;t1_start := FALSE; 
    ELSIF ((x0 = FALSE) AND  (t0.Q = TRUE) AND  (t1.Q = FALSE)) THEN 
        cstate16 := 22643; y0 := FALSE; y1 := FALSE; y2 := FALSE; t0_start := FALSE;t1_start := FALSE; 
    ELSIF ((x0 = FALSE) AND  (t0.Q = TRUE) AND  (t1.Q = TRUE)) THEN 
        cstate16 := 22644; y0 := FALSE; y1 := FALSE; y2 := FALSE; t0_start := FALSE;t1_start := FALSE; 
    ELSIF ((x0 = TRUE) AND  (t0.Q = FALSE) AND  (t1.Q = FALSE)) THEN 
        cstate16 := 26033; y0 := TRUE; y1 := FALSE; y2 := FALSE; t0_start := FALSE;t1_start := FALSE; 
    ELSIF ((x0 = TRUE) AND  (t0.Q = FALSE) AND  (t1.Q = TRUE)) THEN 
        cstate16 := 26034; y0 := TRUE; y1 := FALSE; y2 := FALSE; t0_start := FALSE;t1_start := FALSE; 
    ELSIF ((x0 = TRUE) AND  (t0.Q = TRUE) AND  (t1.Q = FALSE)) THEN 
        cstate16 := 43409; y0 := TRUE; y1 := FALSE; y2 := FALSE; t0_start := FALSE;t1_start := FALSE; 
    ELSIF ((x0 = TRUE) AND  (t0.Q = TRUE) AND  (t1.Q = TRUE)) THEN 
        cstate16 := 43410; y0 := TRUE; y1 := FALSE; y2 := FALSE; t0_start := FALSE;t1_start := FALSE; 
    END_IF;
20673:
    IF ((x0 = FALSE) AND  (t0.Q = FALSE) AND  (t1.Q = FALSE)) THEN 
        cstate16 := 26739; y0 := FALSE; y1 := FALSE; y2 := FALSE; t0_start := FALSE;t1_start := FALSE; 
    ELSIF ((x0 = FALSE) AND  (t0.Q = FALSE) AND  (t1.Q = TRUE)) THEN 
        cstate16 := 26740; y0 := FALSE; y1 := FALSE; y2 := FALSE; t0_start := FALSE;t1_start := FALSE; 
    ELSIF ((x0 = FALSE) AND  (t0.Q = TRUE) AND  (t1.Q = FALSE)) THEN 
        cstate16 := 22643; y0 := FALSE; y1 := FALSE; y2 := FALSE; t0_start := FALSE;t1_start := FALSE; 
    ELSIF ((x0 = FALSE) AND  (t0.Q = TRUE) AND  (t1.Q = TRUE)) THEN 
        cstate16 := 22644; y0 := FALSE; y1 := FALSE; y2 := FALSE; t0_start := FALSE;t1_start := FALSE; 
    ELSIF ((x0 = TRUE) AND  (t0.Q = FALSE) AND  (t1.Q = FALSE)) THEN 
        cstate16 := 26033; y0 := TRUE; y1 := FALSE; y2 := FALSE; t0_start := FALSE;t1_start := FALSE; 
    ELSIF ((x0 = TRUE) AND  (t0.Q = FALSE) AND  (t1.Q = TRUE)) THEN 
        cstate16 := 26038; y0 := TRUE; y1 := FALSE; y2 := TRUE; t0_start := FALSE;t1_start := FALSE; 
    ELSIF ((x0 = TRUE) AND  (t0.Q = TRUE) AND  (t1.Q = FALSE)) THEN 
        cstate16 := 43409; y0 := TRUE; y1 := FALSE; y2 := FALSE; t0_start := FALSE;t1_start := FALSE; 
    ELSIF ((x0 = TRUE) AND  (t0.Q = TRUE) AND  (t1.Q = TRUE)) THEN 
        cstate16 := 43414; y0 := TRUE; y1 := FALSE; y2 := TRUE; t0_start := FALSE;t1_start := FALSE; 
    END_IF;
26034:
    IF ((x0 = FALSE) AND  (t0.Q = FALSE) AND  (t1.Q = FALSE)) THEN 
        cstate16 := 26739; y0 := FALSE; y1 := FALSE; y2 := FALSE; t0_start := FALSE;t1_start := FALSE; 
    ELSIF ((x0 = FALSE) AND  (t0.Q = FALSE) AND  (t1.Q = TRUE)) THEN 
        cstate16 := 26740; y0 := FALSE; y1 := FALSE; y2 := FALSE; t0_start := FALSE;t1_start := FALSE; 
    ELSIF ((x0 = FALSE) AND  (t0.Q = TRUE) AND  (t1.Q = FALSE)) THEN 
        cstate16 := 17491; y0 := FALSE; y1 := FALSE; y2 := FALSE; t0_start := FALSE;t1_start := TRUE; t1_up := FALSE; 
    ELSIF ((x0 = FALSE) AND  (t0.Q = TRUE) AND  (t1.Q = TRUE)) THEN 
        cstate16 := 17492; y0 := FALSE; y1 := FALSE; y2 := FALSE; t0_start := FALSE;t1_start := TRUE; t1_up := FALSE; 
    ELSIF ((x0 = TRUE) AND  (t0.Q = FALSE) AND  (t1.Q = FALSE)) THEN 
        cstate16 := 26033; y0 := TRUE; y1 := FALSE; y2 := FALSE; t0_start := FALSE;t1_start := FALSE; 
    ELSIF ((x0 = TRUE) AND  (t0.Q = FALSE) AND  (t1.Q = TRUE)) THEN 
        cstate16 := 26034; y0 := TRUE; y1 := FALSE; y2 := FALSE; t0_start := FALSE;t1_start := FALSE; 
    ELSIF ((x0 = TRUE) AND  (t0.Q = TRUE) AND  (t1.Q = FALSE)) THEN 
        cstate16 := 42449; y0 := TRUE; y1 := TRUE; y2 := FALSE; t0_start := FALSE;t1_start := TRUE; t1_up := FALSE; 
    ELSIF ((x0 = TRUE) AND  (t0.Q = TRUE) AND  (t1.Q = TRUE)) THEN 
        cstate16 := 42450; y0 := TRUE; y1 := TRUE; y2 := FALSE; t0_start := FALSE;t1_start := TRUE; t1_up := FALSE; 
    END_IF;
26033:
    IF ((x0 = FALSE) AND  (t0.Q = FALSE) AND  (t1.Q = FALSE)) THEN 
        cstate16 := 26739; y0 := FALSE; y1 := FALSE; y2 := FALSE; t0_start := FALSE;t1_start := FALSE; 
    ELSIF ((x0 = FALSE) AND  (t0.Q = FALSE) AND  (t1.Q = TRUE)) THEN 
        cstate16 := 26740; y0 := FALSE; y1 := FALSE; y2 := FALSE; t0_start := FALSE;t1_start := FALSE; 
    ELSIF ((x0 = FALSE) AND  (t0.Q = TRUE) AND  (t1.Q = FALSE)) THEN 
        cstate16 := 17491; y0 := FALSE; y1 := FALSE; y2 := FALSE; t0_start := FALSE;t1_start := TRUE; t1_up := FALSE; 
    ELSIF ((x0 = FALSE) AND  (t0.Q = TRUE) AND  (t1.Q = TRUE)) THEN 
        cstate16 := 17492; y0 := FALSE; y1 := FALSE; y2 := FALSE; t0_start := FALSE;t1_start := TRUE; t1_up := FALSE; 
    ELSIF ((x0 = TRUE) AND  (t0.Q = FALSE) AND  (t1.Q = FALSE)) THEN 
        cstate16 := 26033; y0 := TRUE; y1 := FALSE; y2 := FALSE; t0_start := FALSE;t1_start := FALSE; 
    ELSIF ((x0 = TRUE) AND  (t0.Q = FALSE) AND  (t1.Q = TRUE)) THEN 
        cstate16 := 26038; y0 := TRUE; y1 := FALSE; y2 := TRUE; t0_start := FALSE;t1_start := FALSE; 
    ELSIF ((x0 = TRUE) AND  (t0.Q = TRUE) AND  (t1.Q = FALSE)) THEN 
        cstate16 := 42449; y0 := TRUE; y1 := TRUE; y2 := FALSE; t0_start := FALSE;t1_start := TRUE; t1_up := FALSE; 
    ELSIF ((x0 = TRUE) AND  (t0.Q = TRUE) AND  (t1.Q = TRUE)) THEN 
        cstate16 := 42453; y0 := TRUE; y1 := TRUE; y2 := TRUE; t0_start := FALSE;t1_start := TRUE; t1_up := FALSE; 
    END_IF;
28788:
    IF ((x0 = FALSE) AND  (t0.Q = FALSE) AND  (t1.Q = FALSE)) THEN 
        cstate16 := 34931; y0 := FALSE; y1 := FALSE; y2 := FALSE; t0_start := FALSE;t1_start := FALSE; 
    ELSIF ((x0 = FALSE) AND  (t0.Q = FALSE) AND  (t1.Q = TRUE)) THEN 
        cstate16 := 34932; y0 := FALSE; y1 := FALSE; y2 := FALSE; t0_start := FALSE;t1_start := FALSE; 
    ELSIF ((x0 = FALSE) AND  (t0.Q = TRUE) AND  (t1.Q = FALSE)) THEN 
        cstate16 := 28787; y0 := FALSE; y1 := FALSE; y2 := FALSE; t0_start := FALSE;t1_start := FALSE; 
    ELSIF ((x0 = FALSE) AND  (t0.Q = TRUE) AND  (t1.Q = TRUE)) THEN 
        cstate16 := 28788; y0 := FALSE; y1 := FALSE; y2 := FALSE; t0_start := FALSE;t1_start := FALSE; 
    ELSIF ((x0 = TRUE) AND  (t0.Q = FALSE) AND  (t1.Q = FALSE)) THEN 
        cstate16 := 40163; y0 := TRUE; y1 := FALSE; y2 := FALSE; t0_start := TRUE; t0_up := FALSE;t1_start := FALSE; 
    ELSIF ((x0 = TRUE) AND  (t0.Q = FALSE) AND  (t1.Q = TRUE)) THEN 
        cstate16 := 40164; y0 := TRUE; y1 := FALSE; y2 := FALSE; t0_start := TRUE; t0_up := FALSE;t1_start := FALSE; 
    ELSIF ((x0 = TRUE) AND  (t0.Q = TRUE) AND  (t1.Q = FALSE)) THEN 
        cstate16 := 39139; y0 := TRUE; y1 := FALSE; y2 := FALSE; t0_start := TRUE; t0_up := FALSE;t1_start := FALSE; 
    ELSIF ((x0 = TRUE) AND  (t0.Q = TRUE) AND  (t1.Q = TRUE)) THEN 
        cstate16 := 39140; y0 := TRUE; y1 := FALSE; y2 := FALSE; t0_start := TRUE; t0_up := FALSE;t1_start := FALSE; 
    END_IF;
28787:
    IF ((x0 = FALSE) AND  (t0.Q = FALSE) AND  (t1.Q = FALSE)) THEN 
        cstate16 := 34931; y0 := FALSE; y1 := FALSE; y2 := FALSE; t0_start := FALSE;t1_start := FALSE; 
    ELSIF ((x0 = FALSE) AND  (t0.Q = FALSE) AND  (t1.Q = TRUE)) THEN 
        cstate16 := 34932; y0 := FALSE; y1 := FALSE; y2 := FALSE; t0_start := FALSE;t1_start := FALSE; 
    ELSIF ((x0 = FALSE) AND  (t0.Q = TRUE) AND  (t1.Q = FALSE)) THEN 
        cstate16 := 28787; y0 := FALSE; y1 := FALSE; y2 := FALSE; t0_start := FALSE;t1_start := FALSE; 
    ELSIF ((x0 = FALSE) AND  (t0.Q = TRUE) AND  (t1.Q = TRUE)) THEN 
        cstate16 := 28788; y0 := FALSE; y1 := FALSE; y2 := FALSE; t0_start := FALSE;t1_start := FALSE; 
    ELSIF ((x0 = TRUE) AND  (t0.Q = FALSE) AND  (t1.Q = FALSE)) THEN 
        cstate16 := 40163; y0 := TRUE; y1 := FALSE; y2 := FALSE; t0_start := TRUE; t0_up := FALSE;t1_start := FALSE; 
    ELSIF ((x0 = TRUE) AND  (t0.Q = FALSE) AND  (t1.Q = TRUE)) THEN 
        cstate16 := 40167; y0 := TRUE; y1 := FALSE; y2 := TRUE; t0_start := TRUE; t0_up := FALSE;t1_start := FALSE; 
    ELSIF ((x0 = TRUE) AND  (t0.Q = TRUE) AND  (t1.Q = FALSE)) THEN 
        cstate16 := 39139; y0 := TRUE; y1 := FALSE; y2 := FALSE; t0_start := TRUE; t0_up := FALSE;t1_start := FALSE; 
    ELSIF ((x0 = TRUE) AND  (t0.Q = TRUE) AND  (t1.Q = TRUE)) THEN 
        cstate16 := 39143; y0 := TRUE; y1 := FALSE; y2 := TRUE; t0_start := TRUE; t0_up := FALSE;t1_start := FALSE; 
    END_IF;
40172:
    IF ((x0 = FALSE) AND  (t0.Q = FALSE) AND  (t1.Q = FALSE)) THEN 
        cstate16 := 26739; y0 := FALSE; y1 := FALSE; y2 := FALSE; t0_start := FALSE;t1_start := FALSE; 
    ELSIF ((x0 = FALSE) AND  (t0.Q = FALSE) AND  (t1.Q = TRUE)) THEN 
        cstate16 := 26740; y0 := FALSE; y1 := FALSE; y2 := FALSE; t0_start := FALSE;t1_start := FALSE; 
    ELSIF ((x0 = FALSE) AND  (t0.Q = TRUE) AND  (t1.Q = FALSE)) THEN 
        cstate16 := 17491; y0 := FALSE; y1 := FALSE; y2 := FALSE; t0_start := FALSE;t1_start := TRUE; t1_up := FALSE; 
    ELSIF ((x0 = FALSE) AND  (t0.Q = TRUE) AND  (t1.Q = TRUE)) THEN 
        cstate16 := 17492; y0 := FALSE; y1 := FALSE; y2 := FALSE; t0_start := FALSE;t1_start := TRUE; t1_up := FALSE; 
    ELSIF ((x0 = TRUE) AND  (t0.Q = FALSE) AND  (t1.Q = FALSE)) THEN 
        cstate16 := 40540; y0 := TRUE; y1 := FALSE; y2 := TRUE; t0_start := FALSE;t1_start := FALSE; 
    ELSIF ((x0 = TRUE) AND  (t0.Q = FALSE) AND  (t1.Q = TRUE)) THEN 
        cstate16 := 40535; y0 := TRUE; y1 := FALSE; y2 := TRUE; t0_start := FALSE;t1_start := FALSE; 
    ELSIF ((x0 = TRUE) AND  (t0.Q = TRUE) AND  (t1.Q = FALSE)) THEN 
        cstate16 := 46651; y0 := TRUE; y1 := TRUE; y2 := TRUE; t0_start := FALSE;t1_start := TRUE; t1_up := FALSE; 
    ELSIF ((x0 = TRUE) AND  (t0.Q = TRUE) AND  (t1.Q = TRUE)) THEN 
        cstate16 := 46648; y0 := TRUE; y1 := TRUE; y2 := TRUE; t0_start := FALSE;t1_start := TRUE; t1_up := FALSE; 
    END_IF;
40652:
    IF ((x0 = FALSE) AND  (t0.Q = FALSE) AND  (t1.Q = FALSE)) THEN 
        cstate16 := 26739; y0 := FALSE; y1 := FALSE; y2 := FALSE; t0_start := FALSE;t1_start := FALSE; 
    ELSIF ((x0 = FALSE) AND  (t0.Q = FALSE) AND  (t1.Q = TRUE)) THEN 
        cstate16 := 26740; y0 := FALSE; y1 := FALSE; y2 := FALSE; t0_start := FALSE;t1_start := FALSE; 
    ELSIF ((x0 = FALSE) AND  (t0.Q = TRUE) AND  (t1.Q = FALSE)) THEN 
        cstate16 := 17491; y0 := FALSE; y1 := FALSE; y2 := FALSE; t0_start := FALSE;t1_start := TRUE; t1_up := FALSE; 
    ELSIF ((x0 = FALSE) AND  (t0.Q = TRUE) AND  (t1.Q = TRUE)) THEN 
        cstate16 := 17492; y0 := FALSE; y1 := FALSE; y2 := FALSE; t0_start := FALSE;t1_start := TRUE; t1_up := FALSE; 
    ELSIF ((x0 = TRUE) AND  (t0.Q = FALSE) AND  (t1.Q = FALSE)) THEN 
        cstate16 := 40668; y0 := TRUE; y1 := TRUE; y2 := TRUE; t0_start := FALSE;t1_start := FALSE; 
    ELSIF ((x0 = TRUE) AND  (t0.Q = FALSE) AND  (t1.Q = TRUE)) THEN 
        cstate16 := 40663; y0 := TRUE; y1 := TRUE; y2 := TRUE; t0_start := FALSE;t1_start := FALSE; 
    ELSIF ((x0 = TRUE) AND  (t0.Q = TRUE) AND  (t1.Q = FALSE)) THEN 
        cstate16 := 46651; y0 := TRUE; y1 := TRUE; y2 := TRUE; t0_start := FALSE;t1_start := TRUE; t1_up := FALSE; 
    ELSIF ((x0 = TRUE) AND  (t0.Q = TRUE) AND  (t1.Q = TRUE)) THEN 
        cstate16 := 46648; y0 := TRUE; y1 := TRUE; y2 := TRUE; t0_start := FALSE;t1_start := TRUE; t1_up := FALSE; 
    END_IF;
41635:
    IF ((x0 = FALSE) AND  (t0.Q = FALSE) AND  (t1.Q = FALSE)) THEN 
        cstate16 := 23667; y0 := FALSE; y1 := FALSE; y2 := FALSE; t0_start := FALSE;t1_start := FALSE; 
    ELSIF ((x0 = FALSE) AND  (t0.Q = FALSE) AND  (t1.Q = TRUE)) THEN 
        cstate16 := 26740; y0 := FALSE; y1 := FALSE; y2 := FALSE; t0_start := FALSE;t1_start := FALSE; 
    ELSIF ((x0 = FALSE) AND  (t0.Q = TRUE) AND  (t1.Q = FALSE)) THEN 
        cstate16 := 17491; y0 := FALSE; y1 := FALSE; y2 := FALSE; t0_start := FALSE;t1_start := TRUE; t1_up := FALSE; 
    ELSIF ((x0 = FALSE) AND  (t0.Q = TRUE) AND  (t1.Q = TRUE)) THEN 
        cstate16 := 17492; y0 := FALSE; y1 := FALSE; y2 := FALSE; t0_start := FALSE;t1_start := TRUE; t1_up := FALSE; 
    ELSIF ((x0 = TRUE) AND  (t0.Q = FALSE) AND  (t1.Q = FALSE)) THEN 
        cstate16 := 41699; y0 := TRUE; y1 := TRUE; y2 := FALSE; t0_start := FALSE;t1_start := FALSE; 
    ELSIF ((x0 = TRUE) AND  (t0.Q = FALSE) AND  (t1.Q = TRUE)) THEN 
        cstate16 := 40663; y0 := TRUE; y1 := TRUE; y2 := TRUE; t0_start := FALSE;t1_start := FALSE; 
    ELSIF ((x0 = TRUE) AND  (t0.Q = TRUE) AND  (t1.Q = FALSE)) THEN 
        cstate16 := 46643; y0 := TRUE; y1 := TRUE; y2 := FALSE; t0_start := FALSE;t1_start := TRUE; t1_up := FALSE; 
    ELSIF ((x0 = TRUE) AND  (t0.Q = TRUE) AND  (t1.Q = TRUE)) THEN 
        cstate16 := 46648; y0 := TRUE; y1 := TRUE; y2 := TRUE; t0_start := FALSE;t1_start := TRUE; t1_up := FALSE; 
    END_IF;
40659:
    IF ((x0 = FALSE) AND  (t0.Q = FALSE) AND  (t1.Q = FALSE)) THEN 
        cstate16 := 26739; y0 := FALSE; y1 := FALSE; y2 := FALSE; t0_start := FALSE;t1_start := FALSE; 
    ELSIF ((x0 = FALSE) AND  (t0.Q = FALSE) AND  (t1.Q = TRUE)) THEN 
        cstate16 := 26740; y0 := FALSE; y1 := FALSE; y2 := FALSE; t0_start := FALSE;t1_start := FALSE; 
    ELSIF ((x0 = FALSE) AND  (t0.Q = TRUE) AND  (t1.Q = FALSE)) THEN 
        cstate16 := 17491; y0 := FALSE; y1 := FALSE; y2 := FALSE; t0_start := FALSE;t1_start := TRUE; t1_up := FALSE; 
    ELSIF ((x0 = FALSE) AND  (t0.Q = TRUE) AND  (t1.Q = TRUE)) THEN 
        cstate16 := 17492; y0 := FALSE; y1 := FALSE; y2 := FALSE; t0_start := FALSE;t1_start := TRUE; t1_up := FALSE; 
    ELSIF ((x0 = TRUE) AND  (t0.Q = FALSE) AND  (t1.Q = FALSE)) THEN 
        cstate16 := 40659; y0 := TRUE; y1 := TRUE; y2 := FALSE; t0_start := FALSE;t1_start := FALSE; 
    ELSIF ((x0 = TRUE) AND  (t0.Q = FALSE) AND  (t1.Q = TRUE)) THEN 
        cstate16 := 40663; y0 := TRUE; y1 := TRUE; y2 := TRUE; t0_start := FALSE;t1_start := FALSE; 
    ELSIF ((x0 = TRUE) AND  (t0.Q = TRUE) AND  (t1.Q = FALSE)) THEN 
        cstate16 := 46643; y0 := TRUE; y1 := TRUE; y2 := FALSE; t0_start := FALSE;t1_start := TRUE; t1_up := FALSE; 
    ELSIF ((x0 = TRUE) AND  (t0.Q = TRUE) AND  (t1.Q = TRUE)) THEN 
        cstate16 := 46648; y0 := TRUE; y1 := TRUE; y2 := TRUE; t0_start := FALSE;t1_start := TRUE; t1_up := FALSE; 
    END_IF;
22643:
    IF ((x0 = FALSE) AND  (t0.Q = FALSE) AND  (t1.Q = FALSE)) THEN 
        cstate16 := 34931; y0 := FALSE; y1 := FALSE; y2 := FALSE; t0_start := FALSE;t1_start := FALSE; 
    ELSIF ((x0 = FALSE) AND  (t0.Q = FALSE) AND  (t1.Q = TRUE)) THEN 
        cstate16 := 34932; y0 := FALSE; y1 := FALSE; y2 := FALSE; t0_start := FALSE;t1_start := FALSE; 
    ELSIF ((x0 = FALSE) AND  (t0.Q = TRUE) AND  (t1.Q = FALSE)) THEN 
        cstate16 := 28787; y0 := FALSE; y1 := FALSE; y2 := FALSE; t0_start := FALSE;t1_start := FALSE; 
    ELSIF ((x0 = FALSE) AND  (t0.Q = TRUE) AND  (t1.Q = TRUE)) THEN 
        cstate16 := 28788; y0 := FALSE; y1 := FALSE; y2 := FALSE; t0_start := FALSE;t1_start := FALSE; 
    ELSIF ((x0 = TRUE) AND  (t0.Q = FALSE) AND  (t1.Q = FALSE)) THEN 
        cstate16 := 40163; y0 := TRUE; y1 := FALSE; y2 := FALSE; t0_start := TRUE; t0_up := FALSE;t1_start := FALSE; 
    ELSIF ((x0 = TRUE) AND  (t0.Q = FALSE) AND  (t1.Q = TRUE)) THEN 
        cstate16 := 40167; y0 := TRUE; y1 := FALSE; y2 := TRUE; t0_start := TRUE; t0_up := FALSE;t1_start := FALSE; 
    ELSIF ((x0 = TRUE) AND  (t0.Q = TRUE) AND  (t1.Q = FALSE)) THEN 
        cstate16 := 39139; y0 := TRUE; y1 := FALSE; y2 := FALSE; t0_start := TRUE; t0_up := FALSE;t1_start := FALSE; 
    ELSIF ((x0 = TRUE) AND  (t0.Q = TRUE) AND  (t1.Q = TRUE)) THEN 
        cstate16 := 39143; y0 := TRUE; y1 := FALSE; y2 := TRUE; t0_start := TRUE; t0_up := FALSE;t1_start := FALSE; 
    END_IF;
22644:
    IF ((x0 = FALSE) AND  (t0.Q = FALSE) AND  (t1.Q = FALSE)) THEN 
        cstate16 := 34931; y0 := FALSE; y1 := FALSE; y2 := FALSE; t0_start := FALSE;t1_start := FALSE; 
    ELSIF ((x0 = FALSE) AND  (t0.Q = FALSE) AND  (t1.Q = TRUE)) THEN 
        cstate16 := 34932; y0 := FALSE; y1 := FALSE; y2 := FALSE; t0_start := FALSE;t1_start := FALSE; 
    ELSIF ((x0 = FALSE) AND  (t0.Q = TRUE) AND  (t1.Q = FALSE)) THEN 
        cstate16 := 28787; y0 := FALSE; y1 := FALSE; y2 := FALSE; t0_start := FALSE;t1_start := FALSE; 
    ELSIF ((x0 = FALSE) AND  (t0.Q = TRUE) AND  (t1.Q = TRUE)) THEN 
        cstate16 := 28788; y0 := FALSE; y1 := FALSE; y2 := FALSE; t0_start := FALSE;t1_start := FALSE; 
    ELSIF ((x0 = TRUE) AND  (t0.Q = FALSE) AND  (t1.Q = FALSE)) THEN 
        cstate16 := 40163; y0 := TRUE; y1 := FALSE; y2 := FALSE; t0_start := TRUE; t0_up := FALSE;t1_start := FALSE; 
    ELSIF ((x0 = TRUE) AND  (t0.Q = FALSE) AND  (t1.Q = TRUE)) THEN 
        cstate16 := 40164; y0 := TRUE; y1 := FALSE; y2 := FALSE; t0_start := TRUE; t0_up := FALSE;t1_start := FALSE; 
    ELSIF ((x0 = TRUE) AND  (t0.Q = TRUE) AND  (t1.Q = FALSE)) THEN 
        cstate16 := 39139; y0 := TRUE; y1 := FALSE; y2 := FALSE; t0_start := TRUE; t0_up := FALSE;t1_start := FALSE; 
    ELSIF ((x0 = TRUE) AND  (t0.Q = TRUE) AND  (t1.Q = TRUE)) THEN 
        cstate16 := 39140; y0 := TRUE; y1 := FALSE; y2 := FALSE; t0_start := TRUE; t0_up := FALSE;t1_start := FALSE; 
    END_IF;
8354:
    IF ((x0 = FALSE) AND  (t0.Q = FALSE) AND  (t1.Q = FALSE)) THEN 
        cstate16 := 32883; y0 := FALSE; y1 := FALSE; y2 := FALSE; t0_start := FALSE;t1_start := FALSE; 
    ELSIF ((x0 = FALSE) AND  (t0.Q = FALSE) AND  (t1.Q = TRUE)) THEN 
        cstate16 := 34932; y0 := FALSE; y1 := FALSE; y2 := FALSE; t0_start := FALSE;t1_start := FALSE; 
    ELSIF ((x0 = FALSE) AND  (t0.Q = TRUE) AND  (t1.Q = FALSE)) THEN 
        cstate16 := 27763; y0 := FALSE; y1 := FALSE; y2 := FALSE; t0_start := FALSE;t1_start := FALSE; 
    ELSIF ((x0 = FALSE) AND  (t0.Q = TRUE) AND  (t1.Q = TRUE)) THEN 
        cstate16 := 28788; y0 := FALSE; y1 := FALSE; y2 := FALSE; t0_start := FALSE;t1_start := FALSE; 
    ELSIF ((x0 = TRUE) AND  (t0.Q = FALSE) AND  (t1.Q = FALSE)) THEN 
        cstate16 := 16689; y0 := FALSE; y1 := TRUE; y2 := FALSE; t0_start := FALSE;t1_start := FALSE; 
    ELSIF ((x0 = TRUE) AND  (t0.Q = FALSE) AND  (t1.Q = TRUE)) THEN 
        cstate16 := 14674; y0 := FALSE; y1 := TRUE; y2 := FALSE; t0_start := FALSE;t1_start := FALSE; 
    ELSIF ((x0 = TRUE) AND  (t0.Q = TRUE) AND  (t1.Q = FALSE)) THEN 
        cstate16 := 8497; y0 := FALSE; y1 := TRUE; y2 := FALSE; t0_start := FALSE;t1_start := FALSE; 
    ELSIF ((x0 = TRUE) AND  (t0.Q = TRUE) AND  (t1.Q = TRUE)) THEN 
        cstate16 := 6482; y0 := FALSE; y1 := TRUE; y2 := FALSE; t0_start := FALSE;t1_start := FALSE; 
    END_IF;
2113:
    IF ((x0 = FALSE) AND  (t0.Q = FALSE) AND  (t1.Q = FALSE)) THEN 
        cstate16 := 34931; y0 := FALSE; y1 := FALSE; y2 := FALSE; t0_start := FALSE;t1_start := FALSE; 
    ELSIF ((x0 = FALSE) AND  (t0.Q = FALSE) AND  (t1.Q = TRUE)) THEN 
        cstate16 := 34932; y0 := FALSE; y1 := FALSE; y2 := FALSE; t0_start := FALSE;t1_start := FALSE; 
    ELSIF ((x0 = FALSE) AND  (t0.Q = TRUE) AND  (t1.Q = FALSE)) THEN 
        cstate16 := 28787; y0 := FALSE; y1 := FALSE; y2 := FALSE; t0_start := FALSE;t1_start := FALSE; 
    ELSIF ((x0 = FALSE) AND  (t0.Q = TRUE) AND  (t1.Q = TRUE)) THEN 
        cstate16 := 28788; y0 := FALSE; y1 := FALSE; y2 := FALSE; t0_start := FALSE;t1_start := FALSE; 
    ELSIF ((x0 = TRUE) AND  (t0.Q = FALSE) AND  (t1.Q = FALSE)) THEN 
        cstate16 := 25793; y0 := TRUE; y1 := FALSE; y2 := FALSE; t0_start := TRUE; t0_up := FALSE;t1_start := FALSE; 
    ELSIF ((x0 = TRUE) AND  (t0.Q = FALSE) AND  (t1.Q = TRUE)) THEN 
        cstate16 := 25798; y0 := TRUE; y1 := FALSE; y2 := TRUE; t0_start := TRUE; t0_up := FALSE;t1_start := FALSE; 
    ELSIF ((x0 = TRUE) AND  (t0.Q = TRUE) AND  (t1.Q = FALSE)) THEN 
        cstate16 := 20673; y0 := TRUE; y1 := FALSE; y2 := FALSE; t0_start := TRUE; t0_up := FALSE;t1_start := FALSE; 
    ELSIF ((x0 = TRUE) AND  (t0.Q = TRUE) AND  (t1.Q = TRUE)) THEN 
        cstate16 := 20678; y0 := TRUE; y1 := FALSE; y2 := TRUE; t0_start := TRUE; t0_up := FALSE;t1_start := FALSE; 
    END_IF;
8353:
    IF ((x0 = FALSE) AND  (t0.Q = FALSE) AND  (t1.Q = FALSE)) THEN 
        cstate16 := 32883; y0 := FALSE; y1 := FALSE; y2 := FALSE; t0_start := FALSE;t1_start := FALSE; 
    ELSIF ((x0 = FALSE) AND  (t0.Q = FALSE) AND  (t1.Q = TRUE)) THEN 
        cstate16 := 34932; y0 := FALSE; y1 := FALSE; y2 := FALSE; t0_start := FALSE;t1_start := FALSE; 
    ELSIF ((x0 = FALSE) AND  (t0.Q = TRUE) AND  (t1.Q = FALSE)) THEN 
        cstate16 := 27763; y0 := FALSE; y1 := FALSE; y2 := FALSE; t0_start := FALSE;t1_start := FALSE; 
    ELSIF ((x0 = FALSE) AND  (t0.Q = TRUE) AND  (t1.Q = TRUE)) THEN 
        cstate16 := 28788; y0 := FALSE; y1 := FALSE; y2 := FALSE; t0_start := FALSE;t1_start := FALSE; 
    ELSIF ((x0 = TRUE) AND  (t0.Q = FALSE) AND  (t1.Q = FALSE)) THEN 
        cstate16 := 16689; y0 := FALSE; y1 := TRUE; y2 := FALSE; t0_start := FALSE;t1_start := FALSE; 
    ELSIF ((x0 = TRUE) AND  (t0.Q = FALSE) AND  (t1.Q = TRUE)) THEN 
        cstate16 := 14678; y0 := FALSE; y1 := TRUE; y2 := TRUE; t0_start := FALSE;t1_start := FALSE; 
    ELSIF ((x0 = TRUE) AND  (t0.Q = TRUE) AND  (t1.Q = FALSE)) THEN 
        cstate16 := 8497; y0 := FALSE; y1 := TRUE; y2 := FALSE; t0_start := FALSE;t1_start := FALSE; 
    ELSIF ((x0 = TRUE) AND  (t0.Q = TRUE) AND  (t1.Q = TRUE)) THEN 
        cstate16 := 6486; y0 := FALSE; y1 := TRUE; y2 := TRUE; t0_start := FALSE;t1_start := FALSE; 
    END_IF;
2114:
    IF ((x0 = FALSE) AND  (t0.Q = FALSE) AND  (t1.Q = FALSE)) THEN 
        cstate16 := 34931; y0 := FALSE; y1 := FALSE; y2 := FALSE; t0_start := FALSE;t1_start := FALSE; 
    ELSIF ((x0 = FALSE) AND  (t0.Q = FALSE) AND  (t1.Q = TRUE)) THEN 
        cstate16 := 34932; y0 := FALSE; y1 := FALSE; y2 := FALSE; t0_start := FALSE;t1_start := FALSE; 
    ELSIF ((x0 = FALSE) AND  (t0.Q = TRUE) AND  (t1.Q = FALSE)) THEN 
        cstate16 := 28787; y0 := FALSE; y1 := FALSE; y2 := FALSE; t0_start := FALSE;t1_start := FALSE; 
    ELSIF ((x0 = FALSE) AND  (t0.Q = TRUE) AND  (t1.Q = TRUE)) THEN 
        cstate16 := 28788; y0 := FALSE; y1 := FALSE; y2 := FALSE; t0_start := FALSE;t1_start := FALSE; 
    ELSIF ((x0 = TRUE) AND  (t0.Q = FALSE) AND  (t1.Q = FALSE)) THEN 
        cstate16 := 25793; y0 := TRUE; y1 := FALSE; y2 := FALSE; t0_start := TRUE; t0_up := FALSE;t1_start := FALSE; 
    ELSIF ((x0 = TRUE) AND  (t0.Q = FALSE) AND  (t1.Q = TRUE)) THEN 
        cstate16 := 25794; y0 := TRUE; y1 := FALSE; y2 := FALSE; t0_start := TRUE; t0_up := FALSE;t1_start := FALSE; 
    ELSIF ((x0 = TRUE) AND  (t0.Q = TRUE) AND  (t1.Q = FALSE)) THEN 
        cstate16 := 20673; y0 := TRUE; y1 := FALSE; y2 := FALSE; t0_start := TRUE; t0_up := FALSE;t1_start := FALSE; 
    ELSIF ((x0 = TRUE) AND  (t0.Q = TRUE) AND  (t1.Q = TRUE)) THEN 
        cstate16 := 20674; y0 := TRUE; y1 := FALSE; y2 := FALSE; t0_start := TRUE; t0_up := FALSE;t1_start := FALSE; 
    END_IF;
8357:
    IF ((x0 = FALSE) AND  (t0.Q = FALSE) AND  (t1.Q = FALSE)) THEN 
        cstate16 := 32883; y0 := FALSE; y1 := FALSE; y2 := FALSE; t0_start := FALSE;t1_start := FALSE; 
    ELSIF ((x0 = FALSE) AND  (t0.Q = FALSE) AND  (t1.Q = TRUE)) THEN 
        cstate16 := 34932; y0 := FALSE; y1 := FALSE; y2 := FALSE; t0_start := FALSE;t1_start := FALSE; 
    ELSIF ((x0 = FALSE) AND  (t0.Q = TRUE) AND  (t1.Q = FALSE)) THEN 
        cstate16 := 27763; y0 := FALSE; y1 := FALSE; y2 := FALSE; t0_start := FALSE;t1_start := FALSE; 
    ELSIF ((x0 = FALSE) AND  (t0.Q = TRUE) AND  (t1.Q = TRUE)) THEN 
        cstate16 := 28788; y0 := FALSE; y1 := FALSE; y2 := FALSE; t0_start := FALSE;t1_start := FALSE; 
    ELSIF ((x0 = TRUE) AND  (t0.Q = FALSE) AND  (t1.Q = FALSE)) THEN 
        cstate16 := 16697; y0 := FALSE; y1 := TRUE; y2 := TRUE; t0_start := FALSE;t1_start := FALSE; 
    ELSIF ((x0 = TRUE) AND  (t0.Q = FALSE) AND  (t1.Q = TRUE)) THEN 
        cstate16 := 14678; y0 := FALSE; y1 := TRUE; y2 := TRUE; t0_start := FALSE;t1_start := FALSE; 
    ELSIF ((x0 = TRUE) AND  (t0.Q = TRUE) AND  (t1.Q = FALSE)) THEN 
        cstate16 := 8505; y0 := FALSE; y1 := TRUE; y2 := TRUE; t0_start := FALSE;t1_start := FALSE; 
    ELSIF ((x0 = TRUE) AND  (t0.Q = TRUE) AND  (t1.Q = TRUE)) THEN 
        cstate16 := 6486; y0 := FALSE; y1 := TRUE; y2 := TRUE; t0_start := FALSE;t1_start := FALSE; 
    END_IF;
26042:
    IF ((x0 = FALSE) AND  (t0.Q = FALSE) AND  (t1.Q = FALSE)) THEN 
        cstate16 := 26739; y0 := FALSE; y1 := FALSE; y2 := FALSE; t0_start := FALSE;t1_start := FALSE; 
    ELSIF ((x0 = FALSE) AND  (t0.Q = FALSE) AND  (t1.Q = TRUE)) THEN 
        cstate16 := 26740; y0 := FALSE; y1 := FALSE; y2 := FALSE; t0_start := FALSE;t1_start := FALSE; 
    ELSIF ((x0 = FALSE) AND  (t0.Q = TRUE) AND  (t1.Q = FALSE)) THEN 
        cstate16 := 17491; y0 := FALSE; y1 := FALSE; y2 := FALSE; t0_start := FALSE;t1_start := TRUE; t1_up := FALSE; 
    ELSIF ((x0 = FALSE) AND  (t0.Q = TRUE) AND  (t1.Q = TRUE)) THEN 
        cstate16 := 17492; y0 := FALSE; y1 := FALSE; y2 := FALSE; t0_start := FALSE;t1_start := TRUE; t1_up := FALSE; 
    ELSIF ((x0 = TRUE) AND  (t0.Q = FALSE) AND  (t1.Q = FALSE)) THEN 
        cstate16 := 26042; y0 := TRUE; y1 := FALSE; y2 := TRUE; t0_start := FALSE;t1_start := FALSE; 
    ELSIF ((x0 = TRUE) AND  (t0.Q = FALSE) AND  (t1.Q = TRUE)) THEN 
        cstate16 := 26038; y0 := TRUE; y1 := FALSE; y2 := TRUE; t0_start := FALSE;t1_start := FALSE; 
    ELSIF ((x0 = TRUE) AND  (t0.Q = TRUE) AND  (t1.Q = FALSE)) THEN 
        cstate16 := 42457; y0 := TRUE; y1 := TRUE; y2 := TRUE; t0_start := FALSE;t1_start := TRUE; t1_up := FALSE; 
    ELSIF ((x0 = TRUE) AND  (t0.Q = TRUE) AND  (t1.Q = TRUE)) THEN 
        cstate16 := 42453; y0 := TRUE; y1 := TRUE; y2 := TRUE; t0_start := FALSE;t1_start := TRUE; t1_up := FALSE; 
    END_IF;
40164:
    IF ((x0 = FALSE) AND  (t0.Q = FALSE) AND  (t1.Q = FALSE)) THEN 
        cstate16 := 26739; y0 := FALSE; y1 := FALSE; y2 := FALSE; t0_start := FALSE;t1_start := FALSE; 
    ELSIF ((x0 = FALSE) AND  (t0.Q = FALSE) AND  (t1.Q = TRUE)) THEN 
        cstate16 := 26740; y0 := FALSE; y1 := FALSE; y2 := FALSE; t0_start := FALSE;t1_start := FALSE; 
    ELSIF ((x0 = FALSE) AND  (t0.Q = TRUE) AND  (t1.Q = FALSE)) THEN 
        cstate16 := 17491; y0 := FALSE; y1 := FALSE; y2 := FALSE; t0_start := FALSE;t1_start := TRUE; t1_up := FALSE; 
    ELSIF ((x0 = FALSE) AND  (t0.Q = TRUE) AND  (t1.Q = TRUE)) THEN 
        cstate16 := 17492; y0 := FALSE; y1 := FALSE; y2 := FALSE; t0_start := FALSE;t1_start := TRUE; t1_up := FALSE; 
    ELSIF ((x0 = TRUE) AND  (t0.Q = FALSE) AND  (t1.Q = FALSE)) THEN 
        cstate16 := 40531; y0 := TRUE; y1 := FALSE; y2 := FALSE; t0_start := FALSE;t1_start := FALSE; 
    ELSIF ((x0 = TRUE) AND  (t0.Q = FALSE) AND  (t1.Q = TRUE)) THEN 
        cstate16 := 40532; y0 := TRUE; y1 := FALSE; y2 := FALSE; t0_start := FALSE;t1_start := FALSE; 
    ELSIF ((x0 = TRUE) AND  (t0.Q = TRUE) AND  (t1.Q = FALSE)) THEN 
        cstate16 := 46643; y0 := TRUE; y1 := TRUE; y2 := FALSE; t0_start := FALSE;t1_start := TRUE; t1_up := FALSE; 
    ELSIF ((x0 = TRUE) AND  (t0.Q = TRUE) AND  (t1.Q = TRUE)) THEN 
        cstate16 := 46644; y0 := TRUE; y1 := TRUE; y2 := FALSE; t0_start := FALSE;t1_start := TRUE; t1_up := FALSE; 
    END_IF;
40163:
    IF ((x0 = FALSE) AND  (t0.Q = FALSE) AND  (t1.Q = FALSE)) THEN 
        cstate16 := 26739; y0 := FALSE; y1 := FALSE; y2 := FALSE; t0_start := FALSE;t1_start := FALSE; 
    ELSIF ((x0 = FALSE) AND  (t0.Q = FALSE) AND  (t1.Q = TRUE)) THEN 
        cstate16 := 26740; y0 := FALSE; y1 := FALSE; y2 := FALSE; t0_start := FALSE;t1_start := FALSE; 
    ELSIF ((x0 = FALSE) AND  (t0.Q = TRUE) AND  (t1.Q = FALSE)) THEN 
        cstate16 := 17491; y0 := FALSE; y1 := FALSE; y2 := FALSE; t0_start := FALSE;t1_start := TRUE; t1_up := FALSE; 
    ELSIF ((x0 = FALSE) AND  (t0.Q = TRUE) AND  (t1.Q = TRUE)) THEN 
        cstate16 := 17492; y0 := FALSE; y1 := FALSE; y2 := FALSE; t0_start := FALSE;t1_start := TRUE; t1_up := FALSE; 
    ELSIF ((x0 = TRUE) AND  (t0.Q = FALSE) AND  (t1.Q = FALSE)) THEN 
        cstate16 := 40531; y0 := TRUE; y1 := FALSE; y2 := FALSE; t0_start := FALSE;t1_start := FALSE; 
    ELSIF ((x0 = TRUE) AND  (t0.Q = FALSE) AND  (t1.Q = TRUE)) THEN 
        cstate16 := 40535; y0 := TRUE; y1 := FALSE; y2 := TRUE; t0_start := FALSE;t1_start := FALSE; 
    ELSIF ((x0 = TRUE) AND  (t0.Q = TRUE) AND  (t1.Q = FALSE)) THEN 
        cstate16 := 46643; y0 := TRUE; y1 := TRUE; y2 := FALSE; t0_start := FALSE;t1_start := TRUE; t1_up := FALSE; 
    ELSIF ((x0 = TRUE) AND  (t0.Q = TRUE) AND  (t1.Q = TRUE)) THEN 
        cstate16 := 46648; y0 := TRUE; y1 := TRUE; y2 := TRUE; t0_start := FALSE;t1_start := TRUE; t1_up := FALSE; 
    END_IF;
46739:
    IF ((x0 = FALSE) AND  (t0.Q = FALSE) AND  (t1.Q = FALSE)) THEN 
        cstate16 := 32883; y0 := FALSE; y1 := FALSE; y2 := FALSE; t0_start := FALSE;t1_start := FALSE; 
    ELSIF ((x0 = FALSE) AND  (t0.Q = FALSE) AND  (t1.Q = TRUE)) THEN 
        cstate16 := 34932; y0 := FALSE; y1 := FALSE; y2 := FALSE; t0_start := FALSE;t1_start := FALSE; 
    ELSIF ((x0 = FALSE) AND  (t0.Q = TRUE) AND  (t1.Q = FALSE)) THEN 
        cstate16 := 27763; y0 := FALSE; y1 := FALSE; y2 := FALSE; t0_start := FALSE;t1_start := FALSE; 
    ELSIF ((x0 = FALSE) AND  (t0.Q = TRUE) AND  (t1.Q = TRUE)) THEN 
        cstate16 := 28788; y0 := FALSE; y1 := FALSE; y2 := FALSE; t0_start := FALSE;t1_start := FALSE; 
    ELSIF ((x0 = TRUE) AND  (t0.Q = FALSE) AND  (t1.Q = FALSE)) THEN 
        cstate16 := 41635; y0 := TRUE; y1 := TRUE; y2 := FALSE; t0_start := TRUE; t0_up := FALSE;t1_start := FALSE; 
    ELSIF ((x0 = TRUE) AND  (t0.Q = FALSE) AND  (t1.Q = TRUE)) THEN 
        cstate16 := 40647; y0 := TRUE; y1 := TRUE; y2 := TRUE; t0_start := TRUE; t0_up := FALSE;t1_start := FALSE; 
    ELSIF ((x0 = TRUE) AND  (t0.Q = TRUE) AND  (t1.Q = FALSE)) THEN 
        cstate16 := 46739; y0 := TRUE; y1 := TRUE; y2 := FALSE; t0_start := FALSE;t1_start := FALSE; 
    ELSIF ((x0 = TRUE) AND  (t0.Q = TRUE) AND  (t1.Q = TRUE)) THEN 
        cstate16 := 47799; y0 := TRUE; y1 := TRUE; y2 := TRUE; t0_start := FALSE;t1_start := FALSE; 
    END_IF;
40167:
    IF ((x0 = FALSE) AND  (t0.Q = FALSE) AND  (t1.Q = FALSE)) THEN 
        cstate16 := 26739; y0 := FALSE; y1 := FALSE; y2 := FALSE; t0_start := FALSE;t1_start := FALSE; 
    ELSIF ((x0 = FALSE) AND  (t0.Q = FALSE) AND  (t1.Q = TRUE)) THEN 
        cstate16 := 26740; y0 := FALSE; y1 := FALSE; y2 := FALSE; t0_start := FALSE;t1_start := FALSE; 
    ELSIF ((x0 = FALSE) AND  (t0.Q = TRUE) AND  (t1.Q = FALSE)) THEN 
        cstate16 := 17491; y0 := FALSE; y1 := FALSE; y2 := FALSE; t0_start := FALSE;t1_start := TRUE; t1_up := FALSE; 
    ELSIF ((x0 = FALSE) AND  (t0.Q = TRUE) AND  (t1.Q = TRUE)) THEN 
        cstate16 := 17492; y0 := FALSE; y1 := FALSE; y2 := FALSE; t0_start := FALSE;t1_start := TRUE; t1_up := FALSE; 
    ELSIF ((x0 = TRUE) AND  (t0.Q = FALSE) AND  (t1.Q = FALSE)) THEN 
        cstate16 := 40540; y0 := TRUE; y1 := FALSE; y2 := TRUE; t0_start := FALSE;t1_start := FALSE; 
    ELSIF ((x0 = TRUE) AND  (t0.Q = FALSE) AND  (t1.Q = TRUE)) THEN 
        cstate16 := 40535; y0 := TRUE; y1 := FALSE; y2 := TRUE; t0_start := FALSE;t1_start := FALSE; 
    ELSIF ((x0 = TRUE) AND  (t0.Q = TRUE) AND  (t1.Q = FALSE)) THEN 
        cstate16 := 46651; y0 := TRUE; y1 := TRUE; y2 := TRUE; t0_start := FALSE;t1_start := TRUE; t1_up := FALSE; 
    ELSIF ((x0 = TRUE) AND  (t0.Q = TRUE) AND  (t1.Q = TRUE)) THEN 
        cstate16 := 46648; y0 := TRUE; y1 := TRUE; y2 := TRUE; t0_start := FALSE;t1_start := TRUE; t1_up := FALSE; 
    END_IF;
40647:
    IF ((x0 = FALSE) AND  (t0.Q = FALSE) AND  (t1.Q = FALSE)) THEN 
        cstate16 := 26739; y0 := FALSE; y1 := FALSE; y2 := FALSE; t0_start := FALSE;t1_start := FALSE; 
    ELSIF ((x0 = FALSE) AND  (t0.Q = FALSE) AND  (t1.Q = TRUE)) THEN 
        cstate16 := 26740; y0 := FALSE; y1 := FALSE; y2 := FALSE; t0_start := FALSE;t1_start := FALSE; 
    ELSIF ((x0 = FALSE) AND  (t0.Q = TRUE) AND  (t1.Q = FALSE)) THEN 
        cstate16 := 17491; y0 := FALSE; y1 := FALSE; y2 := FALSE; t0_start := FALSE;t1_start := TRUE; t1_up := FALSE; 
    ELSIF ((x0 = FALSE) AND  (t0.Q = TRUE) AND  (t1.Q = TRUE)) THEN 
        cstate16 := 17492; y0 := FALSE; y1 := FALSE; y2 := FALSE; t0_start := FALSE;t1_start := TRUE; t1_up := FALSE; 
    ELSIF ((x0 = TRUE) AND  (t0.Q = FALSE) AND  (t1.Q = FALSE)) THEN 
        cstate16 := 40668; y0 := TRUE; y1 := TRUE; y2 := TRUE; t0_start := FALSE;t1_start := FALSE; 
    ELSIF ((x0 = TRUE) AND  (t0.Q = FALSE) AND  (t1.Q = TRUE)) THEN 
        cstate16 := 40663; y0 := TRUE; y1 := TRUE; y2 := TRUE; t0_start := FALSE;t1_start := FALSE; 
    ELSIF ((x0 = TRUE) AND  (t0.Q = TRUE) AND  (t1.Q = FALSE)) THEN 
        cstate16 := 46651; y0 := TRUE; y1 := TRUE; y2 := TRUE; t0_start := FALSE;t1_start := TRUE; t1_up := FALSE; 
    ELSIF ((x0 = TRUE) AND  (t0.Q = TRUE) AND  (t1.Q = TRUE)) THEN 
        cstate16 := 46648; y0 := TRUE; y1 := TRUE; y2 := TRUE; t0_start := FALSE;t1_start := TRUE; t1_up := FALSE; 
    END_IF;
41187:
    IF ((x0 = FALSE) AND  (t0.Q = FALSE) AND  (t1.Q = FALSE)) THEN 
        cstate16 := 23667; y0 := FALSE; y1 := FALSE; y2 := FALSE; t0_start := FALSE;t1_start := FALSE; 
    ELSIF ((x0 = FALSE) AND  (t0.Q = FALSE) AND  (t1.Q = TRUE)) THEN 
        cstate16 := 26740; y0 := FALSE; y1 := FALSE; y2 := FALSE; t0_start := FALSE;t1_start := FALSE; 
    ELSIF ((x0 = FALSE) AND  (t0.Q = TRUE) AND  (t1.Q = FALSE)) THEN 
        cstate16 := 17491; y0 := FALSE; y1 := FALSE; y2 := FALSE; t0_start := FALSE;t1_start := TRUE; t1_up := FALSE; 
    ELSIF ((x0 = FALSE) AND  (t0.Q = TRUE) AND  (t1.Q = TRUE)) THEN 
        cstate16 := 17492; y0 := FALSE; y1 := FALSE; y2 := FALSE; t0_start := FALSE;t1_start := TRUE; t1_up := FALSE; 
    ELSIF ((x0 = TRUE) AND  (t0.Q = FALSE) AND  (t1.Q = FALSE)) THEN 
        cstate16 := 41555; y0 := TRUE; y1 := FALSE; y2 := FALSE; t0_start := FALSE;t1_start := FALSE; 
    ELSIF ((x0 = TRUE) AND  (t0.Q = FALSE) AND  (t1.Q = TRUE)) THEN 
        cstate16 := 40535; y0 := TRUE; y1 := FALSE; y2 := TRUE; t0_start := FALSE;t1_start := FALSE; 
    ELSIF ((x0 = TRUE) AND  (t0.Q = TRUE) AND  (t1.Q = FALSE)) THEN 
        cstate16 := 46643; y0 := TRUE; y1 := TRUE; y2 := FALSE; t0_start := FALSE;t1_start := TRUE; t1_up := FALSE; 
    ELSIF ((x0 = TRUE) AND  (t0.Q = TRUE) AND  (t1.Q = TRUE)) THEN 
        cstate16 := 46648; y0 := TRUE; y1 := TRUE; y2 := TRUE; t0_start := FALSE;t1_start := TRUE; t1_up := FALSE; 
    END_IF;
40644:
    IF ((x0 = FALSE) AND  (t0.Q = FALSE) AND  (t1.Q = FALSE)) THEN 
        cstate16 := 26739; y0 := FALSE; y1 := FALSE; y2 := FALSE; t0_start := FALSE;t1_start := FALSE; 
    ELSIF ((x0 = FALSE) AND  (t0.Q = FALSE) AND  (t1.Q = TRUE)) THEN 
        cstate16 := 26740; y0 := FALSE; y1 := FALSE; y2 := FALSE; t0_start := FALSE;t1_start := FALSE; 
    ELSIF ((x0 = FALSE) AND  (t0.Q = TRUE) AND  (t1.Q = FALSE)) THEN 
        cstate16 := 17491; y0 := FALSE; y1 := FALSE; y2 := FALSE; t0_start := FALSE;t1_start := TRUE; t1_up := FALSE; 
    ELSIF ((x0 = FALSE) AND  (t0.Q = TRUE) AND  (t1.Q = TRUE)) THEN 
        cstate16 := 17492; y0 := FALSE; y1 := FALSE; y2 := FALSE; t0_start := FALSE;t1_start := TRUE; t1_up := FALSE; 
    ELSIF ((x0 = TRUE) AND  (t0.Q = FALSE) AND  (t1.Q = FALSE)) THEN 
        cstate16 := 40659; y0 := TRUE; y1 := TRUE; y2 := FALSE; t0_start := FALSE;t1_start := FALSE; 
    ELSIF ((x0 = TRUE) AND  (t0.Q = FALSE) AND  (t1.Q = TRUE)) THEN 
        cstate16 := 40660; y0 := TRUE; y1 := TRUE; y2 := FALSE; t0_start := FALSE;t1_start := FALSE; 
    ELSIF ((x0 = TRUE) AND  (t0.Q = TRUE) AND  (t1.Q = FALSE)) THEN 
        cstate16 := 46643; y0 := TRUE; y1 := TRUE; y2 := FALSE; t0_start := FALSE;t1_start := TRUE; t1_up := FALSE; 
    ELSIF ((x0 = TRUE) AND  (t0.Q = TRUE) AND  (t1.Q = TRUE)) THEN 
        cstate16 := 46644; y0 := TRUE; y1 := TRUE; y2 := FALSE; t0_start := FALSE;t1_start := TRUE; t1_up := FALSE; 
    END_IF;
40643:
    IF ((x0 = FALSE) AND  (t0.Q = FALSE) AND  (t1.Q = FALSE)) THEN 
        cstate16 := 26739; y0 := FALSE; y1 := FALSE; y2 := FALSE; t0_start := FALSE;t1_start := FALSE; 
    ELSIF ((x0 = FALSE) AND  (t0.Q = FALSE) AND  (t1.Q = TRUE)) THEN 
        cstate16 := 26740; y0 := FALSE; y1 := FALSE; y2 := FALSE; t0_start := FALSE;t1_start := FALSE; 
    ELSIF ((x0 = FALSE) AND  (t0.Q = TRUE) AND  (t1.Q = FALSE)) THEN 
        cstate16 := 17491; y0 := FALSE; y1 := FALSE; y2 := FALSE; t0_start := FALSE;t1_start := TRUE; t1_up := FALSE; 
    ELSIF ((x0 = FALSE) AND  (t0.Q = TRUE) AND  (t1.Q = TRUE)) THEN 
        cstate16 := 17492; y0 := FALSE; y1 := FALSE; y2 := FALSE; t0_start := FALSE;t1_start := TRUE; t1_up := FALSE; 
    ELSIF ((x0 = TRUE) AND  (t0.Q = FALSE) AND  (t1.Q = FALSE)) THEN 
        cstate16 := 40659; y0 := TRUE; y1 := TRUE; y2 := FALSE; t0_start := FALSE;t1_start := FALSE; 
    ELSIF ((x0 = TRUE) AND  (t0.Q = FALSE) AND  (t1.Q = TRUE)) THEN 
        cstate16 := 40663; y0 := TRUE; y1 := TRUE; y2 := TRUE; t0_start := FALSE;t1_start := FALSE; 
    ELSIF ((x0 = TRUE) AND  (t0.Q = TRUE) AND  (t1.Q = FALSE)) THEN 
        cstate16 := 46643; y0 := TRUE; y1 := TRUE; y2 := FALSE; t0_start := FALSE;t1_start := TRUE; t1_up := FALSE; 
    ELSIF ((x0 = TRUE) AND  (t0.Q = TRUE) AND  (t1.Q = TRUE)) THEN 
        cstate16 := 46648; y0 := TRUE; y1 := TRUE; y2 := TRUE; t0_start := FALSE;t1_start := TRUE; t1_up := FALSE; 
    END_IF;
27763:
    IF ((x0 = FALSE) AND  (t0.Q = FALSE) AND  (t1.Q = FALSE)) THEN 
        cstate16 := 32883; y0 := FALSE; y1 := FALSE; y2 := FALSE; t0_start := FALSE;t1_start := FALSE; 
    ELSIF ((x0 = FALSE) AND  (t0.Q = FALSE) AND  (t1.Q = TRUE)) THEN 
        cstate16 := 34932; y0 := FALSE; y1 := FALSE; y2 := FALSE; t0_start := FALSE;t1_start := FALSE; 
    ELSIF ((x0 = FALSE) AND  (t0.Q = TRUE) AND  (t1.Q = FALSE)) THEN 
        cstate16 := 27763; y0 := FALSE; y1 := FALSE; y2 := FALSE; t0_start := FALSE;t1_start := FALSE; 
    ELSIF ((x0 = FALSE) AND  (t0.Q = TRUE) AND  (t1.Q = TRUE)) THEN 
        cstate16 := 28788; y0 := FALSE; y1 := FALSE; y2 := FALSE; t0_start := FALSE;t1_start := FALSE; 
    ELSIF ((x0 = TRUE) AND  (t0.Q = FALSE) AND  (t1.Q = FALSE)) THEN 
        cstate16 := 41187; y0 := TRUE; y1 := FALSE; y2 := FALSE; t0_start := TRUE; t0_up := FALSE;t1_start := FALSE; 
    ELSIF ((x0 = TRUE) AND  (t0.Q = FALSE) AND  (t1.Q = TRUE)) THEN 
        cstate16 := 40167; y0 := TRUE; y1 := FALSE; y2 := TRUE; t0_start := TRUE; t0_up := FALSE;t1_start := FALSE; 
    ELSIF ((x0 = TRUE) AND  (t0.Q = TRUE) AND  (t1.Q = FALSE)) THEN 
        cstate16 := 38115; y0 := TRUE; y1 := FALSE; y2 := FALSE; t0_start := TRUE; t0_up := FALSE;t1_start := FALSE; 
    ELSIF ((x0 = TRUE) AND  (t0.Q = TRUE) AND  (t1.Q = TRUE)) THEN 
        cstate16 := 39143; y0 := TRUE; y1 := FALSE; y2 := TRUE; t0_start := TRUE; t0_up := FALSE;t1_start := FALSE; 
    END_IF;
41699:
    IF ((x0 = FALSE) AND  (t0.Q = FALSE) AND  (t1.Q = FALSE)) THEN 
        cstate16 := 23667; y0 := FALSE; y1 := FALSE; y2 := FALSE; t0_start := FALSE;t1_start := FALSE; 
    ELSIF ((x0 = FALSE) AND  (t0.Q = FALSE) AND  (t1.Q = TRUE)) THEN 
        cstate16 := 26740; y0 := FALSE; y1 := FALSE; y2 := FALSE; t0_start := FALSE;t1_start := FALSE; 
    ELSIF ((x0 = FALSE) AND  (t0.Q = TRUE) AND  (t1.Q = FALSE)) THEN 
        cstate16 := 17491; y0 := FALSE; y1 := FALSE; y2 := FALSE; t0_start := FALSE;t1_start := TRUE; t1_up := FALSE; 
    ELSIF ((x0 = FALSE) AND  (t0.Q = TRUE) AND  (t1.Q = TRUE)) THEN 
        cstate16 := 17492; y0 := FALSE; y1 := FALSE; y2 := FALSE; t0_start := FALSE;t1_start := TRUE; t1_up := FALSE; 
    ELSIF ((x0 = TRUE) AND  (t0.Q = FALSE) AND  (t1.Q = FALSE)) THEN 
        cstate16 := 41699; y0 := TRUE; y1 := TRUE; y2 := FALSE; t0_start := FALSE;t1_start := FALSE; 
    ELSIF ((x0 = TRUE) AND  (t0.Q = FALSE) AND  (t1.Q = TRUE)) THEN 
        cstate16 := 40663; y0 := TRUE; y1 := TRUE; y2 := TRUE; t0_start := FALSE;t1_start := FALSE; 
    ELSIF ((x0 = TRUE) AND  (t0.Q = TRUE) AND  (t1.Q = FALSE)) THEN 
        cstate16 := 46643; y0 := TRUE; y1 := TRUE; y2 := FALSE; t0_start := FALSE;t1_start := TRUE; t1_up := FALSE; 
    ELSIF ((x0 = TRUE) AND  (t0.Q = TRUE) AND  (t1.Q = TRUE)) THEN 
        cstate16 := 46648; y0 := TRUE; y1 := TRUE; y2 := TRUE; t0_start := FALSE;t1_start := TRUE; t1_up := FALSE; 
    END_IF;
8505:
    IF ((x0 = FALSE) AND  (t0.Q = FALSE) AND  (t1.Q = FALSE)) THEN 
        cstate16 := 32883; y0 := FALSE; y1 := FALSE; y2 := FALSE; t0_start := FALSE;t1_start := FALSE; 
    ELSIF ((x0 = FALSE) AND  (t0.Q = FALSE) AND  (t1.Q = TRUE)) THEN 
        cstate16 := 34932; y0 := FALSE; y1 := FALSE; y2 := FALSE; t0_start := FALSE;t1_start := FALSE; 
    ELSIF ((x0 = FALSE) AND  (t0.Q = TRUE) AND  (t1.Q = FALSE)) THEN 
        cstate16 := 27763; y0 := FALSE; y1 := FALSE; y2 := FALSE; t0_start := FALSE;t1_start := FALSE; 
    ELSIF ((x0 = FALSE) AND  (t0.Q = TRUE) AND  (t1.Q = TRUE)) THEN 
        cstate16 := 28788; y0 := FALSE; y1 := FALSE; y2 := FALSE; t0_start := FALSE;t1_start := FALSE; 
    ELSIF ((x0 = TRUE) AND  (t0.Q = FALSE) AND  (t1.Q = FALSE)) THEN 
        cstate16 := 16697; y0 := FALSE; y1 := TRUE; y2 := TRUE; t0_start := FALSE;t1_start := FALSE; 
    ELSIF ((x0 = TRUE) AND  (t0.Q = FALSE) AND  (t1.Q = TRUE)) THEN 
        cstate16 := 14678; y0 := FALSE; y1 := TRUE; y2 := TRUE; t0_start := FALSE;t1_start := FALSE; 
    ELSIF ((x0 = TRUE) AND  (t0.Q = TRUE) AND  (t1.Q = FALSE)) THEN 
        cstate16 := 8505; y0 := FALSE; y1 := TRUE; y2 := TRUE; t0_start := FALSE;t1_start := FALSE; 
    ELSIF ((x0 = TRUE) AND  (t0.Q = TRUE) AND  (t1.Q = TRUE)) THEN 
        cstate16 := 6486; y0 := FALSE; y1 := TRUE; y2 := TRUE; t0_start := FALSE;t1_start := FALSE; 
    END_IF;
46747:
    IF ((x0 = FALSE) AND  (t0.Q = FALSE) AND  (t1.Q = FALSE)) THEN 
        cstate16 := 32883; y0 := FALSE; y1 := FALSE; y2 := FALSE; t0_start := FALSE;t1_start := FALSE; 
    ELSIF ((x0 = FALSE) AND  (t0.Q = FALSE) AND  (t1.Q = TRUE)) THEN 
        cstate16 := 34932; y0 := FALSE; y1 := FALSE; y2 := FALSE; t0_start := FALSE;t1_start := FALSE; 
    ELSIF ((x0 = FALSE) AND  (t0.Q = TRUE) AND  (t1.Q = FALSE)) THEN 
        cstate16 := 27763; y0 := FALSE; y1 := FALSE; y2 := FALSE; t0_start := FALSE;t1_start := FALSE; 
    ELSIF ((x0 = FALSE) AND  (t0.Q = TRUE) AND  (t1.Q = TRUE)) THEN 
        cstate16 := 28788; y0 := FALSE; y1 := FALSE; y2 := FALSE; t0_start := FALSE;t1_start := FALSE; 
    ELSIF ((x0 = TRUE) AND  (t0.Q = FALSE) AND  (t1.Q = FALSE)) THEN 
        cstate16 := 41643; y0 := TRUE; y1 := TRUE; y2 := TRUE; t0_start := TRUE; t0_up := FALSE;t1_start := FALSE; 
    ELSIF ((x0 = TRUE) AND  (t0.Q = FALSE) AND  (t1.Q = TRUE)) THEN 
        cstate16 := 40647; y0 := TRUE; y1 := TRUE; y2 := TRUE; t0_start := TRUE; t0_up := FALSE;t1_start := FALSE; 
    ELSIF ((x0 = TRUE) AND  (t0.Q = TRUE) AND  (t1.Q = FALSE)) THEN 
        cstate16 := 46747; y0 := TRUE; y1 := TRUE; y2 := TRUE; t0_start := FALSE;t1_start := FALSE; 
    ELSIF ((x0 = TRUE) AND  (t0.Q = TRUE) AND  (t1.Q = TRUE)) THEN 
        cstate16 := 47799; y0 := TRUE; y1 := TRUE; y2 := TRUE; t0_start := FALSE;t1_start := FALSE; 
    END_IF;
46644:
    IF ((x0 = FALSE) AND  (t0.Q = FALSE) AND  (t1.Q = FALSE)) THEN 
        cstate16 := 32883; y0 := FALSE; y1 := FALSE; y2 := FALSE; t0_start := FALSE;t1_start := FALSE; 
    ELSIF ((x0 = FALSE) AND  (t0.Q = FALSE) AND  (t1.Q = TRUE)) THEN 
        cstate16 := 34932; y0 := FALSE; y1 := FALSE; y2 := FALSE; t0_start := FALSE;t1_start := FALSE; 
    ELSIF ((x0 = FALSE) AND  (t0.Q = TRUE) AND  (t1.Q = FALSE)) THEN 
        cstate16 := 27763; y0 := FALSE; y1 := FALSE; y2 := FALSE; t0_start := FALSE;t1_start := FALSE; 
    ELSIF ((x0 = FALSE) AND  (t0.Q = TRUE) AND  (t1.Q = TRUE)) THEN 
        cstate16 := 28788; y0 := FALSE; y1 := FALSE; y2 := FALSE; t0_start := FALSE;t1_start := FALSE; 
    ELSIF ((x0 = TRUE) AND  (t0.Q = FALSE) AND  (t1.Q = FALSE)) THEN 
        cstate16 := 41635; y0 := TRUE; y1 := TRUE; y2 := FALSE; t0_start := TRUE; t0_up := FALSE;t1_start := FALSE; 
    ELSIF ((x0 = TRUE) AND  (t0.Q = FALSE) AND  (t1.Q = TRUE)) THEN 
        cstate16 := 40644; y0 := TRUE; y1 := TRUE; y2 := FALSE; t0_start := TRUE; t0_up := FALSE;t1_start := FALSE; 
    ELSIF ((x0 = TRUE) AND  (t0.Q = TRUE) AND  (t1.Q = FALSE)) THEN 
        cstate16 := 46739; y0 := TRUE; y1 := TRUE; y2 := FALSE; t0_start := FALSE;t1_start := FALSE; 
    ELSIF ((x0 = TRUE) AND  (t0.Q = TRUE) AND  (t1.Q = TRUE)) THEN 
        cstate16 := 47796; y0 := TRUE; y1 := TRUE; y2 := FALSE; t0_start := FALSE;t1_start := FALSE; 
    END_IF;
47804:
    IF ((x0 = FALSE) AND  (t0.Q = FALSE) AND  (t1.Q = FALSE)) THEN 
        cstate16 := 34931; y0 := FALSE; y1 := FALSE; y2 := FALSE; t0_start := FALSE;t1_start := FALSE; 
    ELSIF ((x0 = FALSE) AND  (t0.Q = FALSE) AND  (t1.Q = TRUE)) THEN 
        cstate16 := 34932; y0 := FALSE; y1 := FALSE; y2 := FALSE; t0_start := FALSE;t1_start := FALSE; 
    ELSIF ((x0 = FALSE) AND  (t0.Q = TRUE) AND  (t1.Q = FALSE)) THEN 
        cstate16 := 28787; y0 := FALSE; y1 := FALSE; y2 := FALSE; t0_start := FALSE;t1_start := FALSE; 
    ELSIF ((x0 = FALSE) AND  (t0.Q = TRUE) AND  (t1.Q = TRUE)) THEN 
        cstate16 := 28788; y0 := FALSE; y1 := FALSE; y2 := FALSE; t0_start := FALSE;t1_start := FALSE; 
    ELSIF ((x0 = TRUE) AND  (t0.Q = FALSE) AND  (t1.Q = FALSE)) THEN 
        cstate16 := 40652; y0 := TRUE; y1 := TRUE; y2 := TRUE; t0_start := TRUE; t0_up := FALSE;t1_start := FALSE; 
    ELSIF ((x0 = TRUE) AND  (t0.Q = FALSE) AND  (t1.Q = TRUE)) THEN 
        cstate16 := 40647; y0 := TRUE; y1 := TRUE; y2 := TRUE; t0_start := TRUE; t0_up := FALSE;t1_start := FALSE; 
    ELSIF ((x0 = TRUE) AND  (t0.Q = TRUE) AND  (t1.Q = FALSE)) THEN 
        cstate16 := 47804; y0 := TRUE; y1 := TRUE; y2 := TRUE; t0_start := FALSE;t1_start := FALSE; 
    ELSIF ((x0 = TRUE) AND  (t0.Q = TRUE) AND  (t1.Q = TRUE)) THEN 
        cstate16 := 47799; y0 := TRUE; y1 := TRUE; y2 := TRUE; t0_start := FALSE;t1_start := FALSE; 
    END_IF;
46643:
    IF ((x0 = FALSE) AND  (t0.Q = FALSE) AND  (t1.Q = FALSE)) THEN 
        cstate16 := 32883; y0 := FALSE; y1 := FALSE; y2 := FALSE; t0_start := FALSE;t1_start := FALSE; 
    ELSIF ((x0 = FALSE) AND  (t0.Q = FALSE) AND  (t1.Q = TRUE)) THEN 
        cstate16 := 34932; y0 := FALSE; y1 := FALSE; y2 := FALSE; t0_start := FALSE;t1_start := FALSE; 
    ELSIF ((x0 = FALSE) AND  (t0.Q = TRUE) AND  (t1.Q = FALSE)) THEN 
        cstate16 := 27763; y0 := FALSE; y1 := FALSE; y2 := FALSE; t0_start := FALSE;t1_start := FALSE; 
    ELSIF ((x0 = FALSE) AND  (t0.Q = TRUE) AND  (t1.Q = TRUE)) THEN 
        cstate16 := 28788; y0 := FALSE; y1 := FALSE; y2 := FALSE; t0_start := FALSE;t1_start := FALSE; 
    ELSIF ((x0 = TRUE) AND  (t0.Q = FALSE) AND  (t1.Q = FALSE)) THEN 
        cstate16 := 41635; y0 := TRUE; y1 := TRUE; y2 := FALSE; t0_start := TRUE; t0_up := FALSE;t1_start := FALSE; 
    ELSIF ((x0 = TRUE) AND  (t0.Q = FALSE) AND  (t1.Q = TRUE)) THEN 
        cstate16 := 40647; y0 := TRUE; y1 := TRUE; y2 := TRUE; t0_start := TRUE; t0_up := FALSE;t1_start := FALSE; 
    ELSIF ((x0 = TRUE) AND  (t0.Q = TRUE) AND  (t1.Q = FALSE)) THEN 
        cstate16 := 46739; y0 := TRUE; y1 := TRUE; y2 := FALSE; t0_start := FALSE;t1_start := FALSE; 
    ELSIF ((x0 = TRUE) AND  (t0.Q = TRUE) AND  (t1.Q = TRUE)) THEN 
        cstate16 := 47799; y0 := TRUE; y1 := TRUE; y2 := TRUE; t0_start := FALSE;t1_start := FALSE; 
    END_IF;
23667:
    IF ((x0 = FALSE) AND  (t0.Q = FALSE) AND  (t1.Q = FALSE)) THEN 
        cstate16 := 23667; y0 := FALSE; y1 := FALSE; y2 := FALSE; t0_start := FALSE;t1_start := FALSE; 
    ELSIF ((x0 = FALSE) AND  (t0.Q = FALSE) AND  (t1.Q = TRUE)) THEN 
        cstate16 := 26740; y0 := FALSE; y1 := FALSE; y2 := FALSE; t0_start := FALSE;t1_start := FALSE; 
    ELSIF ((x0 = FALSE) AND  (t0.Q = TRUE) AND  (t1.Q = FALSE)) THEN 
        cstate16 := 17491; y0 := FALSE; y1 := FALSE; y2 := FALSE; t0_start := FALSE;t1_start := TRUE; t1_up := FALSE; 
    ELSIF ((x0 = FALSE) AND  (t0.Q = TRUE) AND  (t1.Q = TRUE)) THEN 
        cstate16 := 17492; y0 := FALSE; y1 := FALSE; y2 := FALSE; t0_start := FALSE;t1_start := TRUE; t1_up := FALSE; 
    ELSIF ((x0 = TRUE) AND  (t0.Q = FALSE) AND  (t1.Q = FALSE)) THEN 
        cstate16 := 41187; y0 := TRUE; y1 := FALSE; y2 := FALSE; t0_start := TRUE; t0_up := FALSE;t1_start := FALSE; 
    ELSIF ((x0 = TRUE) AND  (t0.Q = FALSE) AND  (t1.Q = TRUE)) THEN 
        cstate16 := 40167; y0 := TRUE; y1 := FALSE; y2 := TRUE; t0_start := TRUE; t0_up := FALSE;t1_start := FALSE; 
    ELSIF ((x0 = TRUE) AND  (t0.Q = TRUE) AND  (t1.Q = FALSE)) THEN 
        cstate16 := 38147; y0 := TRUE; y1 := TRUE; y2 := FALSE; t0_start := TRUE; t0_up := FALSE;t1_start := TRUE; t1_up := FALSE; 
    ELSIF ((x0 = TRUE) AND  (t0.Q = TRUE) AND  (t1.Q = TRUE)) THEN 
        cstate16 := 38152; y0 := TRUE; y1 := TRUE; y2 := TRUE; t0_start := TRUE; t0_up := FALSE;t1_start := TRUE; t1_up := FALSE; 
    END_IF;
19669:
    IF ((x0 = FALSE) AND  (t0.Q = FALSE) AND  (t1.Q = FALSE)) THEN 
        cstate16 := 23667; y0 := FALSE; y1 := FALSE; y2 := FALSE; t0_start := FALSE;t1_start := FALSE; 
    ELSIF ((x0 = FALSE) AND  (t0.Q = FALSE) AND  (t1.Q = TRUE)) THEN 
        cstate16 := 26740; y0 := FALSE; y1 := FALSE; y2 := FALSE; t0_start := FALSE;t1_start := FALSE; 
    ELSIF ((x0 = FALSE) AND  (t0.Q = TRUE) AND  (t1.Q = FALSE)) THEN 
        cstate16 := 17523; y0 := FALSE; y1 := FALSE; y2 := FALSE; t0_start := FALSE;t1_start := FALSE; 
    ELSIF ((x0 = FALSE) AND  (t0.Q = TRUE) AND  (t1.Q = TRUE)) THEN 
        cstate16 := 22644; y0 := FALSE; y1 := FALSE; y2 := FALSE; t0_start := FALSE;t1_start := FALSE; 
    ELSIF ((x0 = TRUE) AND  (t0.Q = FALSE) AND  (t1.Q = FALSE)) THEN 
        cstate16 := 25129; y0 := TRUE; y1 := TRUE; y2 := TRUE; t0_start := FALSE;t1_start := FALSE; 
    ELSIF ((x0 = TRUE) AND  (t0.Q = FALSE) AND  (t1.Q = TRUE)) THEN 
        cstate16 := 26134; y0 := TRUE; y1 := TRUE; y2 := TRUE; t0_start := FALSE;t1_start := FALSE; 
    ELSIF ((x0 = TRUE) AND  (t0.Q = TRUE) AND  (t1.Q = FALSE)) THEN 
        cstate16 := 42489; y0 := TRUE; y1 := TRUE; y2 := TRUE; t0_start := FALSE;t1_start := FALSE; 
    ELSIF ((x0 = TRUE) AND  (t0.Q = TRUE) AND  (t1.Q = TRUE)) THEN 
        cstate16 := 43526; y0 := TRUE; y1 := TRUE; y2 := TRUE; t0_start := FALSE;t1_start := FALSE; 
    END_IF;
16697:
    IF ((x0 = FALSE) AND  (t0.Q = FALSE) AND  (t1.Q = FALSE)) THEN 
        cstate16 := 32883; y0 := FALSE; y1 := FALSE; y2 := FALSE; t0_start := FALSE;t1_start := FALSE; 
    ELSIF ((x0 = FALSE) AND  (t0.Q = FALSE) AND  (t1.Q = TRUE)) THEN 
        cstate16 := 34932; y0 := FALSE; y1 := FALSE; y2 := FALSE; t0_start := FALSE;t1_start := FALSE; 
    ELSIF ((x0 = FALSE) AND  (t0.Q = TRUE) AND  (t1.Q = FALSE)) THEN 
        cstate16 := 27731; y0 := FALSE; y1 := FALSE; y2 := FALSE; t0_start := FALSE;t1_start := TRUE; t1_up := FALSE; 
    ELSIF ((x0 = FALSE) AND  (t0.Q = TRUE) AND  (t1.Q = TRUE)) THEN 
        cstate16 := 27732; y0 := FALSE; y1 := FALSE; y2 := FALSE; t0_start := FALSE;t1_start := TRUE; t1_up := FALSE; 
    ELSIF ((x0 = TRUE) AND  (t0.Q = FALSE) AND  (t1.Q = FALSE)) THEN 
        cstate16 := 16697; y0 := FALSE; y1 := TRUE; y2 := TRUE; t0_start := FALSE;t1_start := FALSE; 
    ELSIF ((x0 = TRUE) AND  (t0.Q = FALSE) AND  (t1.Q = TRUE)) THEN 
        cstate16 := 14678; y0 := FALSE; y1 := TRUE; y2 := TRUE; t0_start := FALSE;t1_start := FALSE; 
    ELSIF ((x0 = TRUE) AND  (t0.Q = TRUE) AND  (t1.Q = FALSE)) THEN 
        cstate16 := 8361; y0 := FALSE; y1 := TRUE; y2 := TRUE; t0_start := FALSE;t1_start := TRUE; t1_up := FALSE; 
    ELSIF ((x0 = TRUE) AND  (t0.Q = TRUE) AND  (t1.Q = TRUE)) THEN 
        cstate16 := 8357; y0 := FALSE; y1 := TRUE; y2 := TRUE; t0_start := FALSE;t1_start := TRUE; t1_up := FALSE; 
    END_IF;
46648:
    IF ((x0 = FALSE) AND  (t0.Q = FALSE) AND  (t1.Q = FALSE)) THEN 
        cstate16 := 32883; y0 := FALSE; y1 := FALSE; y2 := FALSE; t0_start := FALSE;t1_start := FALSE; 
    ELSIF ((x0 = FALSE) AND  (t0.Q = FALSE) AND  (t1.Q = TRUE)) THEN 
        cstate16 := 34932; y0 := FALSE; y1 := FALSE; y2 := FALSE; t0_start := FALSE;t1_start := FALSE; 
    ELSIF ((x0 = FALSE) AND  (t0.Q = TRUE) AND  (t1.Q = FALSE)) THEN 
        cstate16 := 27763; y0 := FALSE; y1 := FALSE; y2 := FALSE; t0_start := FALSE;t1_start := FALSE; 
    ELSIF ((x0 = FALSE) AND  (t0.Q = TRUE) AND  (t1.Q = TRUE)) THEN 
        cstate16 := 28788; y0 := FALSE; y1 := FALSE; y2 := FALSE; t0_start := FALSE;t1_start := FALSE; 
    ELSIF ((x0 = TRUE) AND  (t0.Q = FALSE) AND  (t1.Q = FALSE)) THEN 
        cstate16 := 41643; y0 := TRUE; y1 := TRUE; y2 := TRUE; t0_start := TRUE; t0_up := FALSE;t1_start := FALSE; 
    ELSIF ((x0 = TRUE) AND  (t0.Q = FALSE) AND  (t1.Q = TRUE)) THEN 
        cstate16 := 40647; y0 := TRUE; y1 := TRUE; y2 := TRUE; t0_start := TRUE; t0_up := FALSE;t1_start := FALSE; 
    ELSIF ((x0 = TRUE) AND  (t0.Q = TRUE) AND  (t1.Q = FALSE)) THEN 
        cstate16 := 46747; y0 := TRUE; y1 := TRUE; y2 := TRUE; t0_start := FALSE;t1_start := FALSE; 
    ELSIF ((x0 = TRUE) AND  (t0.Q = TRUE) AND  (t1.Q = TRUE)) THEN 
        cstate16 := 47799; y0 := TRUE; y1 := TRUE; y2 := TRUE; t0_start := FALSE;t1_start := FALSE; 
    END_IF;
39139:
    IF ((x0 = FALSE) AND  (t0.Q = FALSE) AND  (t1.Q = FALSE)) THEN 
        cstate16 := 26739; y0 := FALSE; y1 := FALSE; y2 := FALSE; t0_start := FALSE;t1_start := FALSE; 
    ELSIF ((x0 = FALSE) AND  (t0.Q = FALSE) AND  (t1.Q = TRUE)) THEN 
        cstate16 := 26740; y0 := FALSE; y1 := FALSE; y2 := FALSE; t0_start := FALSE;t1_start := FALSE; 
    ELSIF ((x0 = FALSE) AND  (t0.Q = TRUE) AND  (t1.Q = FALSE)) THEN 
        cstate16 := 22643; y0 := FALSE; y1 := FALSE; y2 := FALSE; t0_start := FALSE;t1_start := FALSE; 
    ELSIF ((x0 = FALSE) AND  (t0.Q = TRUE) AND  (t1.Q = TRUE)) THEN 
        cstate16 := 22644; y0 := FALSE; y1 := FALSE; y2 := FALSE; t0_start := FALSE;t1_start := FALSE; 
    ELSIF ((x0 = TRUE) AND  (t0.Q = FALSE) AND  (t1.Q = FALSE)) THEN 
        cstate16 := 40531; y0 := TRUE; y1 := FALSE; y2 := FALSE; t0_start := FALSE;t1_start := FALSE; 
    ELSIF ((x0 = TRUE) AND  (t0.Q = FALSE) AND  (t1.Q = TRUE)) THEN 
        cstate16 := 40535; y0 := TRUE; y1 := FALSE; y2 := TRUE; t0_start := FALSE;t1_start := FALSE; 
    ELSIF ((x0 = TRUE) AND  (t0.Q = TRUE) AND  (t1.Q = FALSE)) THEN 
        cstate16 := 47683; y0 := TRUE; y1 := FALSE; y2 := FALSE; t0_start := FALSE;t1_start := FALSE; 
    ELSIF ((x0 = TRUE) AND  (t0.Q = TRUE) AND  (t1.Q = TRUE)) THEN 
        cstate16 := 47687; y0 := TRUE; y1 := FALSE; y2 := TRUE; t0_start := FALSE;t1_start := FALSE; 
    END_IF;
19665:
    IF ((x0 = FALSE) AND  (t0.Q = FALSE) AND  (t1.Q = FALSE)) THEN 
        cstate16 := 23667; y0 := FALSE; y1 := FALSE; y2 := FALSE; t0_start := FALSE;t1_start := FALSE; 
    ELSIF ((x0 = FALSE) AND  (t0.Q = FALSE) AND  (t1.Q = TRUE)) THEN 
        cstate16 := 26740; y0 := FALSE; y1 := FALSE; y2 := FALSE; t0_start := FALSE;t1_start := FALSE; 
    ELSIF ((x0 = FALSE) AND  (t0.Q = TRUE) AND  (t1.Q = FALSE)) THEN 
        cstate16 := 17523; y0 := FALSE; y1 := FALSE; y2 := FALSE; t0_start := FALSE;t1_start := FALSE; 
    ELSIF ((x0 = FALSE) AND  (t0.Q = TRUE) AND  (t1.Q = TRUE)) THEN 
        cstate16 := 22644; y0 := FALSE; y1 := FALSE; y2 := FALSE; t0_start := FALSE;t1_start := FALSE; 
    ELSIF ((x0 = TRUE) AND  (t0.Q = FALSE) AND  (t1.Q = FALSE)) THEN 
        cstate16 := 25121; y0 := TRUE; y1 := TRUE; y2 := FALSE; t0_start := FALSE;t1_start := FALSE; 
    ELSIF ((x0 = TRUE) AND  (t0.Q = FALSE) AND  (t1.Q = TRUE)) THEN 
        cstate16 := 26134; y0 := TRUE; y1 := TRUE; y2 := TRUE; t0_start := FALSE;t1_start := FALSE; 
    ELSIF ((x0 = TRUE) AND  (t0.Q = TRUE) AND  (t1.Q = FALSE)) THEN 
        cstate16 := 42481; y0 := TRUE; y1 := TRUE; y2 := FALSE; t0_start := FALSE;t1_start := FALSE; 
    ELSIF ((x0 = TRUE) AND  (t0.Q = TRUE) AND  (t1.Q = TRUE)) THEN 
        cstate16 := 43526; y0 := TRUE; y1 := TRUE; y2 := TRUE; t0_start := FALSE;t1_start := FALSE; 
    END_IF;
19666:
    IF ((x0 = FALSE) AND  (t0.Q = FALSE) AND  (t1.Q = FALSE)) THEN 
        cstate16 := 23667; y0 := FALSE; y1 := FALSE; y2 := FALSE; t0_start := FALSE;t1_start := FALSE; 
    ELSIF ((x0 = FALSE) AND  (t0.Q = FALSE) AND  (t1.Q = TRUE)) THEN 
        cstate16 := 26740; y0 := FALSE; y1 := FALSE; y2 := FALSE; t0_start := FALSE;t1_start := FALSE; 
    ELSIF ((x0 = FALSE) AND  (t0.Q = TRUE) AND  (t1.Q = FALSE)) THEN 
        cstate16 := 17523; y0 := FALSE; y1 := FALSE; y2 := FALSE; t0_start := FALSE;t1_start := FALSE; 
    ELSIF ((x0 = FALSE) AND  (t0.Q = TRUE) AND  (t1.Q = TRUE)) THEN 
        cstate16 := 22644; y0 := FALSE; y1 := FALSE; y2 := FALSE; t0_start := FALSE;t1_start := FALSE; 
    ELSIF ((x0 = TRUE) AND  (t0.Q = FALSE) AND  (t1.Q = FALSE)) THEN 
        cstate16 := 25121; y0 := TRUE; y1 := TRUE; y2 := FALSE; t0_start := FALSE;t1_start := FALSE; 
    ELSIF ((x0 = TRUE) AND  (t0.Q = FALSE) AND  (t1.Q = TRUE)) THEN 
        cstate16 := 26130; y0 := TRUE; y1 := TRUE; y2 := FALSE; t0_start := FALSE;t1_start := FALSE; 
    ELSIF ((x0 = TRUE) AND  (t0.Q = TRUE) AND  (t1.Q = FALSE)) THEN 
        cstate16 := 42481; y0 := TRUE; y1 := TRUE; y2 := FALSE; t0_start := FALSE;t1_start := FALSE; 
    ELSIF ((x0 = TRUE) AND  (t0.Q = TRUE) AND  (t1.Q = TRUE)) THEN 
        cstate16 := 43522; y0 := TRUE; y1 := TRUE; y2 := FALSE; t0_start := FALSE;t1_start := FALSE; 
    END_IF;
38152:
    IF ((x0 = FALSE) AND  (t0.Q = FALSE) AND  (t1.Q = FALSE)) THEN 
        cstate16 := 23667; y0 := FALSE; y1 := FALSE; y2 := FALSE; t0_start := FALSE;t1_start := FALSE; 
    ELSIF ((x0 = FALSE) AND  (t0.Q = FALSE) AND  (t1.Q = TRUE)) THEN 
        cstate16 := 26740; y0 := FALSE; y1 := FALSE; y2 := FALSE; t0_start := FALSE;t1_start := FALSE; 
    ELSIF ((x0 = FALSE) AND  (t0.Q = TRUE) AND  (t1.Q = FALSE)) THEN 
        cstate16 := 17523; y0 := FALSE; y1 := FALSE; y2 := FALSE; t0_start := FALSE;t1_start := FALSE; 
    ELSIF ((x0 = FALSE) AND  (t0.Q = TRUE) AND  (t1.Q = TRUE)) THEN 
        cstate16 := 22644; y0 := FALSE; y1 := FALSE; y2 := FALSE; t0_start := FALSE;t1_start := FALSE; 
    ELSIF ((x0 = TRUE) AND  (t0.Q = FALSE) AND  (t1.Q = FALSE)) THEN 
        cstate16 := 41707; y0 := TRUE; y1 := TRUE; y2 := TRUE; t0_start := FALSE;t1_start := FALSE; 
    ELSIF ((x0 = TRUE) AND  (t0.Q = FALSE) AND  (t1.Q = TRUE)) THEN 
        cstate16 := 40663; y0 := TRUE; y1 := TRUE; y2 := TRUE; t0_start := FALSE;t1_start := FALSE; 
    ELSIF ((x0 = TRUE) AND  (t0.Q = TRUE) AND  (t1.Q = FALSE)) THEN 
        cstate16 := 46747; y0 := TRUE; y1 := TRUE; y2 := TRUE; t0_start := FALSE;t1_start := FALSE; 
    ELSIF ((x0 = TRUE) AND  (t0.Q = TRUE) AND  (t1.Q = TRUE)) THEN 
        cstate16 := 47799; y0 := TRUE; y1 := TRUE; y2 := TRUE; t0_start := FALSE;t1_start := FALSE; 
    END_IF;
END_CASE;

(* Additional processing to handle clocks - in CODESYS, it only starts
    with rising edge and can not be placed inside IF statement *) 
IF(t0_up = TRUE) THEN
    t0_reset := TRUE;
ELSIF(t0_start = TRUE AND t0_up = FALSE) THEN
    t0_up := TRUE;  t0_reset := FALSE;
END_IF
t0(IN:=t0_reset, PT:=T0_VALUE); 
IF(t1_up = TRUE) THEN
    t1_reset := TRUE;
ELSIF(t1_start = TRUE AND t1_up = FALSE) THEN
    t1_up := TRUE;  t1_reset := FALSE;
END_IF
t1(IN:=t1_reset, PT:=T1_VALUE);

END_FUNCTION_BLOCK
